  STRUCT
   GRAPHIC_INIT : BOOL ;	//NEW FL Graphic Init
   EMERGENCY_BLINK : BOOL ;	//NEW FL Emergency Blink
   ON_SW : BOOL ;	//NEW FLS On Sw Temporary
   COMPRESSED_AIR : BOOL ;	//NEW FLS Compressed Air
   AERIAL_LINK_RUN_PB : BOOL ;	//NEW FLS 508 Link Run SW - Diabled
   PACKET_in_FLIPPER_SW : BOOL ;	//NEW FLS Service Enable Switch - Disabled
   SERVICE_INIT_PB : BOOL ;	//NEW FLS Service Initialisation PB
   ALL_SERVICE_ENABLE_SW : BOOL ;	//NEW FLS All Services Enable Switch
   SERVICE_SW_1_STATUS : BOOL ;	//NEW FLS Service 1 Switch
   SERVICE_SW_2_STATUS : BOOL ;	//NEW FLS Service 2 Switch
   SERVICE_SW_3_STATUS : BOOL ;	//NEW FLS Service 3 Switch
   SERVICE_SW_1_2_STATUS : BOOL ;	//NEW FLS Service 1 or 2 Switch
   BIT12 : BOOL ;	//NEW FLS Spare
   BIT13 : BOOL ;	//NEW FLS Spare
   SERVICE_SW_2_TIME_ADJ : BOOL ;	//NEW FLS Service 2 Switch - Time Adjust
   PACKETIZER_GATE_STATUS : BOOL ;	//NEW FLS 2145 Packetizer Flap Gate - Status Bit
   E_STOP_CONSOLE_STATUS : BOOL ;	//NEW FL E-Stop Console
   E_STOP_ELEVATOR_STATUS : BOOL ;	//NEW FL E-Stop Elevator
   E_STOP_FLIPPER_STATUS : BOOL ;	//NEW FL E-Stop Flipper
   E_STOP_LOADER_STATUS : BOOL ;	//NEW FL E-Stop Loader
   HAND_FEED_ARROW_STATUS : BOOL ;	//NEW FL Hand Feed Arrow
   ELEVATOR_DOOR_STATUS : BOOL ;	//NEW FL Elevator Door
   FLIPPER_DOOR_STATUS : BOOL ;	//NEW FL Flipper Door
   LOADER_DOOR_STATUS : BOOL ;	//NEW FL Loader Door
   LIGHT_BARRIER_1_STATUS : BOOL ;	//NEW FL Light Barrier 1 - B5.4 Conveyor 1 Exit - Status Bit
   LIGHT_BARRIER_2_STATUS : BOOL ;	//NEW FL Light Barrier 2 - B5.5 Conveyor 2 InFeed - Status Bit
   LIGHT_BARRIER_3_STATUS : BOOL ;	//NEW FL Light Barrier 3 - B6.0 Conveyor 2 Presence - Status Bit
   LIGHT_BARRIER_4_STATUS : BOOL ;	//NEW FL Light Barrier 4 - B6.1 Conveyor 2 Exit - Status Bit
   LIGHT_BARRIER_5_STATUS : BOOL ;	//NEW FL Light Barrier 5 - B6.2 Conveyor 3 InFeed - Status Bit
   LIGHT_BARRIER_6_STATUS : BOOL ;	//NEW FL Light Barrier 6 - B6.4 Conveyor 3 Exit - Status Bit
   LIGHT_BARRIER_B_STATUS : BOOL ;	//NEW FL Light Barrier B - B5.2 Elevator Limit - Status Bit
   LIGHT_BARRIER_A_STATUS : BOOL ;	//NEW FL Light Barrier A - B5.1 Elevator InFeed - Status Bit
   BIT32 : BOOL ;	//NEW FL Pusher 0 Motion
   BIT33 : BOOL ;	//NEW FL Pusher 0 Motion
   BIT34 : BOOL ;	//NEW FL Pusher 0 Motion
   BIT35 : BOOL ;	//NEW FL Pusher 0 Motion
   BIT36 : BOOL ;	//NEW FL Pusher 0 Motion
   BIT37 : BOOL ;	//NEW FL Pusher 0 Motion
   BIT38 : BOOL ;	//NEW FL Pusher 0 Motion
   BIT39 : BOOL ;	//NEW FL Pusher 0 Motion
   BIT40 : BOOL ;	//NEW FL Elevator Motion
   BIT41 : BOOL ;	//NEW FL Elevator Motion
   BIT42 : BOOL ;	//NEW FL Elevator Motion
   BIT43 : BOOL ;	//NEW FL Elevator Motion
   BIT44 : BOOL ;	//NEW FL Elevator Motion
   BIT45 : BOOL ;	//NEW FL Elevator Motion
   BIT46 : BOOL ;	//NEW FL Elevator Motion
   BIT47 : BOOL ;	//NEW FL Elevator Motion
   BIT48 : BOOL ;	//NEW FL Pusher 1 Motion
   BIT49 : BOOL ;	//NEW FL Pusher 1 Motion
   BIT50 : BOOL ;	//NEW FL Pusher 1 Motion
   BIT51 : BOOL ;	//NEW FL Pusher 1 Motion
   BIT52 : BOOL ;	//NEW FL Pusher 1 Motion
   BIT53 : BOOL ;	//NEW FL Pusher 1 Motion
   BIT54 : BOOL ;	//NEW FL Pusher 1 Motion
   BIT55 : BOOL ;	//NEW FL Pusher 1 Motion
   BIT56 : BOOL ;	//NEW FL Pusher 2 Motion
   BIT57 : BOOL ;	//NEW FL Pusher 2 Motion
   BIT58 : BOOL ;	//NEW FL Pusher 2 Motion
   BIT59 : BOOL ;	//NEW FL Pusher 2 Motion
   BIT60 : BOOL ;	//NEW FL Pusher 2 Motion
   BIT61 : BOOL ;	//NEW FL Pusher 2 Motion
   BIT62 : BOOL ;	//NEW FL Pusher 2 Motion
   CONVEYORS_CLEARING : BOOL ;	//NEW FL Conveyors Clearing
   ELEVATOR_MOTOR_STATUS : BOOL ;	//NEW FL Elevator - Motor M42.0 Status Bit
   PUSHER_1_MOTOR_STATUS : BOOL ;	//NEW FL Pusher 1 - Motor M42.6 Status Bit
   CONVEYOR_1_MOTOR_STATUS : BOOL ;	//NEW FL Conv 1 - Motor M43.0 Status Bit
   CONVEYOR_2B_MOTOR_STATUS : BOOL ;	//NEW FL Conv 2 Belt - Motor M43.4 Status Bit
   CONVEYOR_2R_MOTOR_STATUS : BOOL ;	//NEW FL Conv 2 Roller - Motor M43.5 Status Bit
   CONVEYOR_3_MOTOR_STATUS : BOOL ;	//NEW FL Conveyor 3 - Motor M44.0 Status Bit
   CONVEYOR_4_MOTOR_STATUS : BOOL ;	//NEW FL Conveyor 4 - Motor M44.3 Status Bit
   CONVEYOR_5_MOTOR_STATUS : BOOL ;	//NEW FL Conveyor 5 - Motor M45.0 Status Bit
   CONVEYOR_6_MOTOR_STATUS : BOOL ;	//NEW FL Conveyor 6 - Motor M45.3 Status Bit
   CONVEYOR_7_MOTOR_STATUS : BOOL ;	//NEW FL Conveyor 7 - Motor M45.6 Status Bit
   FLIPPER_MOTOR_STATUS : BOOL ;	//NEW FL Flipper Flip - Motor M46.0 Status Bit
   CONVEYOR_8_MOTOR_STATUS : BOOL ;	//NEW FL Conveyor 8 - Motor M46.4 Status Bit
   TURNTABLE_MOTOR_STATUS : BOOL ;	//NEW FL TurnTable - Motor M47.0 Status Bit
   CONVEYOR_9_MOTOR_STATUS : BOOL ;	//NEW FL Conveyor 9 - Motor M47.5 Status Bit
   PUSHER_2_MOTOR_STATUS : BOOL ;	//NEW FL Pusher 2 - Motor M47.6 Status Bit
   CONVEYOR_10_MOTOR_STATUS : BOOL ;	//NEW FL Conveyor 10 - Motor M48.0 Status Bit
   CONVEYOR_11_MOTOR_STATUS : BOOL ;	//NEW FL Conveyor 11 - Motor M48.3 Status Bit
   CONVEYOR_12_MOTOR_STATUS : BOOL ;	//NEW FL Conveyor 12 - Motor M48.6 Status Bit
   CONVEYOR_13_MOTOR_STATUS : BOOL ;	//NEW FL Conveyor 13 - Motor M49.0 Status Bit
   CONVEYOR_21_MOTOR_STATUS : BOOL ;	//NEW FL Conveyor 21 - Motor M53.2 Status Bit
   CONVEYOR_22_MOTOR_STATUS : BOOL ;	//NEW FL Conveyor 22 - Motor M53.4 Status Bit
   CONVEYOR_23_MOTOR_STATUS : BOOL ;	//NEW FL Conveyor 23 - Motor M54.0 Status Bit
   LOADER_LIFT_MOTOR_STATUS : BOOL ;	//NEW FL Loader Lift - Motor M50.0 Status Bit
   LOADER_FING_MOTOR_STATUS : BOOL ;	//NEW FL Loader Fingers - Motor M50.5 Status Bit
   LOADER_BELT_MOTOR_STATUS : BOOL ;	//NEW FL Loader Belt - Motor M51.0 Status Bit
   LIGHT_BARRIER_7_STATUS : BOOL ;	//NEW FL Light Barrier 7 - B6.7 Conv 4 InFeed Sens - Status
   LIGHT_BARRIER_8_STATUS : BOOL ;	//NEW FL Light Barrier 8 - B7.0 Conv 4 Exit Sens - Status
   LIGHT_BARRIER_9_STATUS : BOOL ;	//NEW FL Light Barrier 9 - B7.1 Conv 5 Exit Sens - Status
   LIGHT_BARRIER_10_STATUS : BOOL ;	//NEW FL Light Barrier 10 - B7.2 Conv 6 Slow Sens - Status Bit
   LIGHT_BARRIER_11_STATUS : BOOL ;	//NEW FL Light Barrier 11 - B7.3 Conv 6 Exit Sens - Status Bit
   LIGHT_BARRIER_12_STATUS : BOOL ;	//NEW FL Light Barrier 12 - B7.4 FLipper InFeed Sens - Status Bit
   LIGHT_BARRIER_13_STATUS : BOOL ;	//NEW FL Light Barrier 13 - B8.2 Flipper Exit Sens - Status Bit
   LIGHT_BARRIER_14_STATUS : BOOL ;	//NEW FL Light Barrier 14 - B9.6 Conv 9 InFeed Sens - Status Bit
   LIGHT_BARRIER_15_STATUS : BOOL ;	//NEW FL Light Barrier 15 - B9.7 Conv 9 Packet Sens - Status Bit
   LIGHT_BARRIER_16_STATUS : BOOL ;	//NEW FL Light Barrier 16 - B10.3 Conv 10 Start Sens - Status Bit
   LIGHT_BARRIER_17_STATUS : BOOL ;	//NEW FL Light Barrier 17 - B10.4 Conv 10 InFeed Sens - Status Bit
   LIGHT_BARRIER_18_STATUS : BOOL ;	//NEW FL Light Barrier 18 - B10.5 Conv 10 Full Sens - Status Bit
   LIGHT_BARRIER_19_STATUS : BOOL ;	//NEW FL Light Barrier 19 - B10.6 Conv 10 Exit Sens - Status Bit
   LIGHT_BARRIER_20_STATUS : BOOL ;	//NEW FL Light Barrier 20 - B10.7 Conv 11 Exit Sens - Status Bit
   LIGHT_BARRIER_21_STATUS : BOOL ;	//NEW FL Light Barrier 21 - B11.0 Conv 12 Exit Sens - Status Bit- Status Bit
   LIGHT_BARRIER_22_STATUS : BOOL ;	//NEW FL Light Barrier 22 - B11.1 Conv 13 Slow Sens - Status Bit
   LIGHT_BARRIER_23_STATUS : BOOL ;	//NEW FL Light Barrier 23 - B11.2 Conv 13 Exit Sens - Status Bit
   LIGHT_BARRIER_24_STATUS : BOOL ;	//NEW FL Light Barrier 24 - B12.3 Fingers Delivery Sens - Status Bit
   LIGHT_BARRIER_25_STATUS : BOOL ;	//NEW FL Light Barrier 25 - B13.0 Loader Empty Sens - Status Bit
   LIGHT_BARRIER_26_STATUS : BOOL ;	//NEW FL Light Barrier 26 - B15.4 Conv 21 Exit Sens - Status Bit
   LIGHT_BARRIER_27_STATUS : BOOL ;	//NEW FL Light Barrier 27 - B15.5 Conv 22 Exit Sens - Status Bit
   LIGHT_BARRIER_28_STATUS : BOOL ;	//NEW FL Light Barrier 28 - B15.6 Conv 23 Slow Sens - Status Bit
   LIGHT_BARRIER_29_STATUS : BOOL ;	//NEW FL Light Barrier 29 - B15.7 Conv 23 Exit Sens - Status Bit
   LIGHT_BARRIER_30_STATUS : BOOL ;	//NEW FL Light Barrier 30 - B35.2 Conv 0 InFeed Sens - Status Bit
   LIGHT_BARRIER_31_STATUS : BOOL ;	//NEW FL Light Barrier 31 - B35.3 Conv 0 Exit Sens - Status Bit
   LIGHT_BARRIER_32_STATUS : BOOL ;	//NEW FL Light Barrier 32 - B35.4 Conv 0 Length Sens - Status Bit
   PROX_9_STATUS : BOOL ;	//NEW FL Prox 9 - P8.5 TurnTable Rotation InFeed Slow - Status Bit
   PROX_10_STATUS : BOOL ;	//NEW FL Prox 10 - P8.6 TurnTable Rotation InFeed Stop - Status Bit
   PROX_11_STATUS : BOOL ;	//NEW FL Prox 11 - P9.2 TurnTable Rotation Exit Slow - Status Bit
   PROX_12_STATUS : BOOL ;	//NEW FL Prox 12 - P9.3 TurnTable Rotation Exit Stop - Status Bit
   PROX_13_STATUS : BOOL ;	//NEW FL Prox 13 - P10.0 Pusher 2 Retract Sens - Status Bit
   PROX_14_STATUS : BOOL ;	//NEW FL Prox 14 - P10.1 Pusher 2 Extend Sens - Status Bit
   PROX_15_STATUS : BOOL ;	//NEW FL Prox 15 - P15.0 Pivot 10 High Sens - Status Bit
   PROX_16_STATUS : BOOL ;	//NEW FL Prox 16 - P15.1 Pivot 10 Low Sens - Status Bit
   PROX_17_STATUS : BOOL ;	//NEW FL Prox 17 - P13.2 Loader H Level Stop - Status Bit
   PROX_18_STATUS : BOOL ;	//NEW FL Prox 18 - P13.1 Loader H Level Slow - Status Bit
   PROX_19_STATUS : BOOL ;	//NEW FL Prox 19 - P11.4 Loader L Level Stop - Status Bit
   PROX_20_STATUS : BOOL ;	//NEW FL Prox 20 - P11.5 Loader L Level Slow - Status Bit
   PROX_21_STATUS : BOOL ;	//NEW FL Prox 21 - P11.6 Loader Slow Bot - Status Bit
   PROX_22_STATUS : BOOL ;	//NEW FL Prox 22 - P11.7 Loader Stop Bot - Status Bit
   PROX_23_STATUS : BOOL ;	//NEW FL Prox 23 - P12.0 Loader Finger Retract - Status Bit
   PROX_24_STATUS : BOOL ;	//NEW FL Prox 24 - P12.1 Loader Finger Extend - Status Bit
   FP131 : BOOL ;	//NEW FP One Shot
   FP132 : BOOL ;	//NEW FP One Shot
   FP133 : BOOL ;	//NEW FP One Shot
   FP134 : BOOL ;	//NEW FP One Shot
   FP135 : BOOL ;	//NEW FP One Shot
   TURNTABLE_DELIV_POSITION : BOOL ;	//NEW FL TurnTable Delivery Position
   TURNTABLE_REVERSE_ARROW : BOOL ;	//NEW FL TurnTable Arrow Reverse Packet
   TURNTABLE_DIR_SELECT_SW : BOOL ;	//NEW FL TurnTable Direction Select SW
   TURNTABLE_FLICK_MOTION : BOOL ;	//NEW FL TurnTable Flicker - Motion
   FP140 : BOOL ;	//NEW FP One Shot
   FP141 : BOOL ;	//NEW FP One Shot
   FP142 : BOOL ;	//NEW FP One Shot
   FP143 : BOOL ;	//NEW FP One Shot
   PROX_1_STATUS : BOOL ;	//NEW FL Prox 1 - P4.0 Elevator Bottom Position - Status Bit
   PROX_2_STATUS : BOOL ;	//NEW FL Prox 2 - P4.1 Elevator SlowDown Bot - Status Bit
   PROX_3_STATUS : BOOL ;	//NEW FL Prox 3 - P4.2 Elevator SlowDown Top - Status Bit
   PROX_4_STATUS : BOOL ;	//NEW FL Prox 4 - P4.3 Elevator Top Position - Status Bit
   PROX_5_STATUS : BOOL ;	//NEW FL Prox 5 - P4.4 Pusher 1 Home - Status Bit
   PROX_6_STATUS : BOOL ;	//NEW FL Prox 6 - P4.5 Pusher 1 Limit - Status Bit
   PROX_7_STATUS : BOOL ;	//NEW FL Prox 7 - P8.0 Flipper Fingers Right Position - Status Bit
   PROX_8_STATUS : BOOL ;	//NEW FL Prox 8 - P8.1 Flipper Fingers Left Position - Status Bit
   BIT152 : BOOL ;	//NEW FL Loader Motion
   BIT153 : BOOL ;	//NEW FL Loader Motion
   BIT154 : BOOL ;	//NEW FL Loader Motion
   BIT155 : BOOL ;	//NEW FL Loader Motion
   BIT156 : BOOL ;	//NEW FL Loader Motion
   BIT157 : BOOL ;	//NEW FL Loader Motion
   BIT158 : BOOL ;	//NEW FL Loader Motion
   BIT159 : BOOL ;	//NEW FL Loader Motion
   SERVICE_SSW_MAIN : BOOL ;	//NEW FL Service SW Main Screen
   SERVICE_SSW_STATUS : BOOL ;	//NEW FL Service SW Main Screen - Status
   CLEARING_SSW_MAIN : BOOL ;	//NEW FL Clearing SW Main Screen
   CLEARING_SSW_STATUS : BOOL ;	//NEW FL Clearing SW Main Screen - Status
   MAN_FEED_SSW_MAIN : BOOL ;	//NEW FL Hand Feed SW Main Screen
   MAN_FEED_SSW_STATUS : BOOL ;	//NEW FL Hand Feed SW Main Screen - Status
   TURNTABLE_SSW_MAIN : BOOL ;	//NEW FL Turn Table Turn SW = 1:CCW - 0:CW Main Screen
   TURNTABLE_SSW_STATUS : BOOL ;	//NEW FL Turn Table Select Main Screen - Status
   FLIPPER_SSW_MAIN : BOOL ;	//NEW FL Flipper SW Main Screen
   FLIPPER_SSW_STATUS : BOOL ;	//NEW FL Flipper SW Main Screen - Status
   ROLLER_SSW_MAIN : BOOL ;	//NEW FL Roller SW Main Screen
   ROLLER_SSW_STATUS : BOOL ;	//NEW FL Roller SW Main Screen - Status
   ELEVATOR_ROUND_TRIP_SSW : BOOL ;	//NEW FL Elevator - Round Trip PB
   BIT173 : BOOL ;
   BIT174 : BOOL ;
   BIT175 : BOOL ;
   HMI_PUSHER_0_TEST_SSW : BOOL ;	//NEW FL Pusher 0 SW
   HMI_ELEVATOR_SERVICE_SSW : BOOL ;	//NEW FL Elevator Service SW
   HMI_ELEVATOR_TEST_DN_SSW : BOOL ;	//NEW FL Elevator DN PB
   HMI_ELEVATOR_TEST_UP_SSW : BOOL ;	//NEW FL Elevator UP PB
   HMI_ROLLER_TEST_FWD_SSW : BOOL ;	//NEW FL Roller FWD SW
   HMI_ROLLER_TEST_REV_SSW : BOOL ;	//NEW FL Roller REV SW
   HMI_PUSHER_1_TEST_SSW : BOOL ;	//NEW FL Pusher 1 SW
   HMI_CONVEYOR_1_TEST_SSW : BOOL ;	//NEW FL Conv 1 SW
   HMI_CONVEYOR_2B_TEST_SSW : BOOL ;	//NEW FL Conv 2 Belt SW
   HMI_CONVEYOR_2L_TEST_SSW : BOOL ;	//NEW FL Conv 2 Lift SW
   HMI_CONVEYOR_2R_TEST_SSW : BOOL ;	//NEW FL Conv 2 Roller SW
   HMI_CONVEYOR_3_TEST_SSW : BOOL ;	//NEW FL Conv 3 SW
   HMI_CONVEYOR_4_TEST_SSW : BOOL ;	//NEW FL Conv 4 SW
   HMI_CONVEYOR_5_TEST_SSW : BOOL ;	//NEW FL Conv 5 SW
   HMI_CONVEYOR_6_TEST_SSW : BOOL ;	//NEW FL Conv 6 SW
   HMI_CONVEYOR_7_TEST_SSW : BOOL ;	//NEW FL Flipper Conv 7 SW
   HMI_CONVEYOR_8_TEST_SSW : BOOL ;	//NEW FL Turn Table Conv 8 SW
   HMI_TURNTABLE_CCW_SSW : BOOL ;	//NEW FL Turn Table / Conveyor CCW PB
   HMI_TURNTABLE_CW_SSW : BOOL ;	//NEW FL Turn Table / Conveyor CW PB
   HMI_FLIPPER_SERVICE_SSW : BOOL ;	//NEW FL Flipper Service SW
   HMI_FLIPPER_FLIP_SSW : BOOL ;	//NEW FL Flipper - Flip PB
   HMI_CONVEYOR_9_TEST_SSW : BOOL ;	//NEW FL Conv 9 SW
   HMI_PUSHER_2_TEST_SSW : BOOL ;	//NEW FL Pusher 2 SW
   HMI_PIVOT_SERVICE_SSW : BOOL ;	//NEW FL Conv 10 - Pivot Service SW
   HMI_PIVOT_TEST_DN_SSW : BOOL ;	//NEW FL Conv 10 - Pivot DN PB
   HMI_PIVOT_TEST_UP_SSW : BOOL ;	//NEW FL Conv 10 - Pivot UP PB
   BIT202 : BOOL ;	//NEW FL Spare
   BIT203 : BOOL ;	//NEW FL Spare
   TURNTABLE_SERVICE_PBSHOW : BOOL ;	//NEW FL TurnTable Service PB SHOW
   TURNTABLE_SERVICE_SSW : BOOL ;	//NEW FL TurnTable Service SW
   HMI_CONVEYOR_10_TEST_SSW : BOOL ;	//NEW FL Conv 10 - Conveyor SW
   LOADER_FING_SERVICE_SSW : BOOL ;	//NEW FL Loader Service SW - Fingers
   LOADER_LIFT_SERVICE_SSW : BOOL ;	//NEW FL Loader Service SW - Lift
   LOADER_LIFT_TOP_PB : BOOL ;	//NEW FL Loader Lift - TOP PB
   LOADER_LIFT_UP_PB : BOOL ;	//NEW FL Loader Lift - UP PB
   LOADER_LIFT_DN_PB : BOOL ;	//NEW FL Loader Lift - DOWN PB
   FINGER_RETRACT_TEST_PB : BOOL ;	//NEW FL Loader Fingers Retract PB
   FINGER_EXTEND_TEST_PB : BOOL ;	//NEW FL Loader Fingers Extend PB
   FINGER_TILT_TEST_PB : BOOL ;	//NEW FL Loader Fingers Tilt Down PB
   FINGER_BELT_TEST_SW : BOOL ;	//NEW FL Loader Fingers Belt SW
   HMI_CONVEYOR_11_TEST_SSW : BOOL ;	//NEW FL Conv 11 Test SW
   HMI_CONVEYOR_12_TEST_SSW : BOOL ;	//NEW FL Conv 12 Test SW
   HMI_CONVEYOR_13_TEST_SSW : BOOL ;	//NEW FL Conv 13 Test SW
   HMI_CONVEYOR_21_TEST_SSW : BOOL ;	//NEW FL Conv 21 Test SW
   HMI_CONVEYOR_22_TEST_SSW : BOOL ;	//NEW FL Conv 22 Test SW
   HMI_CONVEYOR_23_TEST_SSW : BOOL ;	//NEW FL Conv 23 Test SW
   CONVEYOR_0_MOTOR_STATUS : BOOL ;	//NEW FL Conveyor 0 - Motor M62.0 Status Bit
   PUSHER_0_MOTOR_STATUS : BOOL ;	//NEW FL Pusher 0 - Motor M62.2 Status Bit
   PUSHER_0_COLOR_WORD : WORD ;	//NEW WD Pusher 0 - 2145 - Motor Status Color
   CONV_0_COLOR_WORD : WORD ;	//NEW WD Conveyor 0 - 2145 - Motor Status Color
   ELEVATOR_COLOR_WORD : WORD ;	//NEW WD Elevator - Motor Status Color
   PUSHER_1_COLOR_WORD : WORD ;	//NEW WD Pusher 1 - Motor Status Color
   CONV_1_COLOR_WORD : WORD ;	//NEW WD Conv 1 - Motor Status Color
   CONV_2_BELT_COLOR_WORD : WORD ;	//NEW WD Conv 2 Belt - Motor Status Color
   LIFT_ROLLER_2_COLOR_WORD : WORD ;	//NEW WD Lift 2 Roller - Actuator Status Color
   CONV_2_ROLLER_COLOR_WORD : WORD ;	//NEW WD Conv 2 Roller - Motor Status Color
   CONV_3_COLOR_WORD : WORD ;	//NEW WD Conveyor 3 - Motor Status Color
   CONV_4_COLOR_WORD : WORD ;	//NEW WD Conveyor 4 - Motor Status Color
   CONV_5_COLOR_WORD : WORD ;	//NEW WD Conveyor 5 - Motor Status Color
   CONV_6_COLOR_WORD : WORD ;	//NEW WD Conveyor 6 - Motor Status Color
   CONV_7_COLOR_WORD : WORD ;	//NEW WD Conveyor 7 - Motor Status Color
   FLIPPER_COLOR_WORD : WORD ;	//NEW WD Flipper - Motor M46.0 Status Color
   CONV_8_COLOR_WORD : WORD ;	//NEW WD Conveyor 8 - Motor M46.4 Status Color
   TURN_TABLE_COLOR_WORD : WORD ;	//NEW WD TurnTable - Motor M47.0 Status Color
   CONV_9_COLOR_WORD : WORD ;	//NEW WD Conveyor 9 - Motor M47.5 Status Color
   PUSHER_2_COLOR_WORD : WORD ;	//NEW WD Pusher 2 - Motor M47.6 Status Color
   CONV_10_COLOR_WORD : WORD ;	//NEW WD Conveyor 10 - Motor M48.0 Status Color
   CONV_11_COLOR_WORD : WORD ;	//NEW WD Conveyor 11 - Motor M48.3 Status Color
   CONV_12_COLOR_WORD : WORD ;	//NEW WD Conveyor 12 - Motor M48.6 Status Color
   CONV_13_COLOR_WORD : WORD ;	//NEW WD Conveyor 13 - Motor M49.0 Status Color
   CONV_21_COLOR_WORD : WORD ;	//NEW WD Conveyor 21 - Motor M53.4 Status Color
   CONV_22_COLOR_WORD : WORD ;	//NEW WD Conveyor 22 - Motor M53.6 Status Color
   CONV_23_COLOR_WORD : WORD ;	//NEW WD Conveyor 23 - Motor M54.0 Status Color
   LOADER_LIFT_COLOR_WORD : WORD ;	//NEW WD Loader Lift - Motor M54.6 Status Color
   LOADER_FING_COLOR_WORD : WORD ;	//NEW WD Loader Fingers - Motor M50.5 Status Color
   FINGERS_BELT_COLOR_WORD : WORD ;	//NEW WD Fingers Belt - Motor M54.6 Status Color
   HIGH_LEVEL_23_GRAPHIC : WORD ;	//NEW WD High Level Conveyor 23
   LOW_LEVEL_13_GRAPHIC : WORD ;	//NEW WD Low Level Conveyor 13
   PIVOT_GRAPHIC : WORD ;	//NEW WD Pivot Conveyor Graphic
   CONV_3_COUNT : WORD ;	//NEW WD Slat Conveyor 3 - Packet Count
   CONV_4_COUNT : WORD ;	//NEW WD Collator Conveyor 4 - Packet Count
   CONV_5_COUNT : WORD ;	//NEW WD Link Conveyor 5 - Packet Count
   CONV_6_COUNT : WORD ;	//NEW WD Delivery Conveyor 6 - Packet Count
   CONV_10_COUNT : WORD ;	//NEW WD Pivot Conveyor 10 - Packet Count
   CONV_11_COUNT : WORD ;	//NEW WD Cumul Conveyor 11 - Packet Count
   CONV_12_COUNT : WORD ;	//NEW WD Cumul Conveyor 12 - Packet Count
   CONV_13_COUNT : WORD ;	//NEW WD Delivery Conveyor 13 - Packet Count
   CONV_21_COUNT : WORD ;	//NEW WD Cumul Conveyor 21 - Packet Count
   CONV_22_COUNT : WORD ;	//NEW WD Cumul Conveyor 22 - Packet Count
   CONV_23_COUNT : WORD ;	//NEW WD Delivery Conveyor 23 - Packet Count
   FLIPPER_CCW : WORD ;	//NEW WD Flipper Graphic CCW
   FLIPPER_CW : WORD ;	//NEW WD Flipper Graphic CW
   FLIPPER_POSITION : WORD ;	//NEW WD Flipper Positioning mS
   TURN_COLOR : WORD ;	//NEW WD Turn Table - Turn Color
   FLIPPER_COLOR : WORD ;	//NEW WD Flipper Color
   FLIPPER_PACK_PRESENCE : WORD ;	//NEW WD Flipper - Packet Presence
   TURNTABLE_PACK_PRESENCE : WORD ;	//NEW WD TurnTable - Packet Presence
   ROLLER_PACK_PRESENCE : WORD ;	//NEW WD Pusher Roller - Packet Presence
   PUSHER_PACK_PRESENCE : WORD ;	//NEW WD Pusher - Packet Presence
   CONV_0_STATUS : BOOL ;	//NEW FL Conveyor 0 - Motor Status Bit
   PUSHER_0_STATUS : BOOL ;	//NEW FL Pusher 0 - Motor Status
   ELEVATOR_STATUS : BOOL ;	//NEW FL Elevator - Motor Status
   PUSHER_1_STATUS : BOOL ;	//NEW FL Pusher 1 - Motor Status
   CONV_1_STATUS : BOOL ;	//NEW FL Conveyor 1 - Motor Status
   TURNTABLE_RNDTRIP : BOOL ;	//NEW FL TurnTable Round Trip CMD
   RNDTRIP_PB_VISIBLE : BOOL ;	//NEW FL TurnTable Round Trip PB Visible
   BOOL_SPARE227 : BOOL ;	//NEW FL
   SCREEN_CALL_0 : BOOL ;	//NEW FL  HMI Call Screen 0
   SCREEN_CALL_1 : BOOL ;	//NEW FL  HMI Call Screen 1
   SCREEN_CALL_2 : BOOL ;	//NEW FL  HMI Call Screen 2
   SCREEN_CALL_3 : BOOL ;	//NEW FL  HMI Call Screen 3
   SCREEN_CALL_4 : BOOL ;	//NEW FL  HMI Call Screen 4
   BOOL_SPARE2276 : BOOL ;	//NEW FL
   BOOL_SPARE2277 : BOOL ;	//NEW FL
   BOOL_SPARE2278 : BOOL ;	//NEW FL
   BOOL_SPARE2279 : BOOL ;	//NEW FL
   BOOL_SPARE22710 : BOOL ;	//NEW FL
   BOOL_SPARE22711 : BOOL ;	//NEW FL
   BOOL_SPARE22712 : BOOL ;	//NEW FL
   BOOL_SPARE22713 : BOOL ;	//NEW FL
   BOOL_SPARE22714 : BOOL ;	//NEW FL
   BOOL_SPARE22715 : BOOL ;	//NEW FL
   BOOL_SPARE22716 : BOOL ;	//NEW FL
   BOOL_SPARE22717 : BOOL ;	//NEW FL
   BOOL_SPARE22718 : BOOL ;	//NEW FL
   BOOL_SPARE22719 : BOOL ;	//NEW FL
   BOOL_SPARE22720 : BOOL ;	//NEW FL
   BOOL_SPARE22721 : BOOL ;	//NEW FL
   BOOL_SPARE22722 : BOOL ;	//NEW FL
   BOOL_SPARE22723 : BOOL ;	//NEW FL
   BOOL_SPARE22724 : BOOL ;	//NEW FL
   WORD_SPARE23 : WORD ;	//NEW WD
   FLIPPER_TURN_COLOR : WORD ;	//NEW WD Flipper Turn Color
   NEW_ORDER_COLOR : WORD ;	//NEW WD Conveyor 10 - New Order Color
   SERVICE_FLIPPER : BOOL ;	//NEW FLS Flipper Service - Switch
   FLIP_TEST : BOOL ;	//NEW FLS Flipper Flip - Test Switch
   SERVICE_TURNTABLE : BOOL ;	//NEW FLS TurnTable Service - Switch
   TURN_TEST_CW : BOOL ;	//NEW FLS TurnTable - Turn CW - Status Bit
   TURN_TEST_CCW : BOOL ;	//NEW FLS TurnTable - Turn CCW - Status Bit
   PUSHER_2_TEST : BOOL ;	//NEW FLS Pusher 2 - Test Switch
   CONVEYOR_10_TEST_SW : BOOL ;	//NEW FLS Collator Conveyor 10 - Test Switch
   PIVOT_SERVICE_SW : BOOL ;	//NEW FL Pivot Service - Status
   PIVOT_UP_TEST_PB : BOOL ;	//NEW FLS Pivot Conveyor UP - Test Switch
   PIVOT_DN_TEST_PB : BOOL ;	//NEW FLS Pivot Conveyor DN - Test Switch
   PIVOT_STATUS : BOOL ;	//NEW FL Pivot ON - Status
   CONV_8_INVERT_SELECT : BOOL ;	//NEW FL TurnTable Conveyor 8 - Positioning Time - Display Selector Bit - INVERT
   CONVEYOR_11_TEST_SW : BOOL ;	//NEW FLS Cumul Conveyor 11 - Test Switch
   CONVEYOR_12_TEST_SW : BOOL ;	//NEW FLS Cumul Conveyor 12 - Test Switch
   CONVEYOR_13_TEST_SW : BOOL ;	//NEW FLS Delivery Conveyor 13 - Test Switch
   CONVEYOR_21_TEST_SW : BOOL ;	//NEW FLS Cumul Conveyor 21 - Test Switch
   CONVEYOR_22_TEST_SW : BOOL ;	//NEW FLS Cumul Conveyor 22 - Test Switch
   CONVEYOR_23_TEST_SW : BOOL ;	//NEW FLS Delivery Conveyor 23 - Test Switch
   LOADER_SERVICE_SW : BOOL ;	//NEW FLS Loader Service - Switch
   LOADER_UP_TEST_PB : BOOL ;	//NEW FLS Loader Lift Up - Test Switch
   LOADER_DN_TEST_PB : BOOL ;	//NEW FLS Loader Lift Dn - Test Switch
   FINGERS_EXTEND_TEST_PB : BOOL ;	//NEW FLS Loader Finger Extend - Test Switch
   FINGERS_RETRACT_TEST_PB : BOOL ;	//NEW FLS Loader Finger Retract - Test Switch
   FP_ONESHOT_0 : BOOL ;	//NEW FP One Shot
   CONVEYOR_0_SERVICE_SW : BOOL ;	//NEW FL Conveyor 0 / Pusher 0 - Service Enable
   ELEVATOR_SERVICE_SW : BOOL ;	//NEW FL Elevator / Pusher 1 - Service Enable
   CONVEYOR_1_SERVICE_SW : BOOL ;	//NEW FL Conveyor 1 - Service Enable Select - Screen 4
   CONVEYOR_2_SERVICE_SW : BOOL ;	//NEW FL Conveyor 2 - Service Enable Select - Screen 4
   CONVEYOR_3_SERVICE_SW : BOOL ;	//NEW FL Conveyor 3 - Service Enable Select - Screen 4
   CONVEYOR_4_SERVICE_SW : BOOL ;	//NEW FL Conveyor 4 - Service Enable Select - Screen 4
   CONVEYOR_5_SERVICE_SW : BOOL ;	//NEW FL Conveyor 5 - Service Enable Select - Screen 4
   CONVEYOR_6_SERVICE_SW : BOOL ;	//NEW FL Conveyor 6 - Service Enable Select - Screen 4
   CONVEYOR_7_SERVICE_SW : BOOL ;	//NEW FL Conveyor 7 / Flipper - Service Enable Select - Screen 4
   CONVEYOR_8_SERVICE_SW : BOOL ;	//NEW FL Conveyor 8 / TurnTable - Service Enable Select - Screen 4
   CONVEYOR_9_SERVICE_SW : BOOL ;	//NEW FL Conveyor 9 / Pusher 2 - Service Enable Select - Screen 4
   CONVEYOR_10_SERVICE_SW : BOOL ;	//NEW FL Conveyor 10 - Service Enable Select - Screen 4
   CONVEYOR_11_SERVICE_SW : BOOL ;	//NEW FL Conveyors 11, 12, 13 - Service Enable Select - Screen 4
   CONVEYOR_21_SERVICE_SW : BOOL ;	//NEW FL Conveyors 21, 22, 23 - Service Enable Select - Screen 4
   LOADER_SERVICE_ENABLE_SW : BOOL ;	//NEW FL Loader - Service Enable
   CTRL48 : BOOL ;	//NEW FL Spare - Service Enable
   CTRL49 : BOOL ;	//NEW FL Spare -
   CTRL50 : BOOL ;	//NEW FL Spare -
   CTRL51 : BOOL ;	//NEW FL Spare -
   CTRL52 : BOOL ;	//NEW FL Spare -
   CTRL53 : BOOL ;	//NEW FL Spare -
   CTRL54 : BOOL ;	//NEW FL Spare -
   CTRL55 : BOOL ;	//NEW FL Spare -
   CTRL56 : BOOL ;	//NEW FL Spare -
   CLEARING_FUNCTION : WORD ;	//NEW WD Clearing Function - Underneat Rectangle
   WORD57 : WORD ;	//NEW WD
   WORD58 : WORD ;	//NEW WD
   ACTUAL_HMI_SCREEN_NO : WORD ;	//NEW WD HMI Actual Display Screen
   CONVEYOR_MAXCOUNT_L : WORD  := W#16#6;	//NEW WD All Conveyors Max Count Lenght (6)
   CONVEYOR_MAXCOUNT_W : WORD  := W#16#7;	//NEW WD All Conveyors Max Count Widtht (7)
   WORD62 : WORD ;	//NEW WD
   CONV_7_POS_mS : WORD ;	//NEW WD Flipper Conveyor 7 - Positioning Time x10 [mS]
   CONV_8_POS_FWD_mS : WORD ;	//NEW WD TurnTable Conveyor 8 - FWD Positioning Time x10 [mS]
   CONV_8_POS_REV_mS : WORD ;	//NEW WD TurnTable Conveyor 8 - REV Positioning Time x10 [mS]
   CONV_9_POS_mS : WORD ;	//NEW WD Pusher 2 Conveyor 9 - Positioning Time x10 [mS]
   WORD_PACKET_LENGTH : WORD ;	//NEW WD Actual Packet Length mm
   DELAY_DISPLAY_7 : WORD ;	//NEW WD HMI Flipper 7 Delay Display
   DELAY_DISPLAY_9 : WORD ;	//NEW WD HMI Conveyor 9 Delay Display
   WORD_SPARE2 : WORD ;
   WORD_SPARE3 : WORD ;
   WORD_SPARE4 : WORD ;
  END_STRUCT ;
BEGIN
   GRAPHIC_INIT := FALSE;
   EMERGENCY_BLINK := FALSE;
   ON_SW := FALSE;
   COMPRESSED_AIR := FALSE;
   AERIAL_LINK_RUN_PB := FALSE;
   PACKET_in_FLIPPER_SW := FALSE;
   SERVICE_INIT_PB := FALSE;
   ALL_SERVICE_ENABLE_SW := FALSE;
   SERVICE_SW_1_STATUS := FALSE;
   SERVICE_SW_2_STATUS := FALSE;
   SERVICE_SW_3_STATUS := FALSE;
   SERVICE_SW_1_2_STATUS := FALSE;
   BIT12 := FALSE;
   BIT13 := FALSE;
   SERVICE_SW_2_TIME_ADJ := FALSE;
   PACKETIZER_GATE_STATUS := FALSE;
   E_STOP_CONSOLE_STATUS := FALSE;
   E_STOP_ELEVATOR_STATUS := FALSE;
   E_STOP_FLIPPER_STATUS := FALSE;
   E_STOP_LOADER_STATUS := FALSE;
   HAND_FEED_ARROW_STATUS := FALSE;
   ELEVATOR_DOOR_STATUS := FALSE;
   FLIPPER_DOOR_STATUS := FALSE;
   LOADER_DOOR_STATUS := FALSE;
   LIGHT_BARRIER_1_STATUS := FALSE;
   LIGHT_BARRIER_2_STATUS := FALSE;
   LIGHT_BARRIER_3_STATUS := FALSE;
   LIGHT_BARRIER_4_STATUS := FALSE;
   LIGHT_BARRIER_5_STATUS := FALSE;
   LIGHT_BARRIER_6_STATUS := FALSE;
   LIGHT_BARRIER_B_STATUS := FALSE;
   LIGHT_BARRIER_A_STATUS := FALSE;
   BIT32 := FALSE;
   BIT33 := FALSE;
   BIT34 := FALSE;
   BIT35 := FALSE;
   BIT36 := FALSE;
   BIT37 := FALSE;
   BIT38 := FALSE;
   BIT39 := FALSE;
   BIT40 := FALSE;
   BIT41 := FALSE;
   BIT42 := FALSE;
   BIT43 := FALSE;
   BIT44 := FALSE;
   BIT45 := FALSE;
   BIT46 := FALSE;
   BIT47 := FALSE;
   BIT48 := FALSE;
   BIT49 := FALSE;
   BIT50 := FALSE;
   BIT51 := FALSE;
   BIT52 := FALSE;
   BIT53 := FALSE;
   BIT54 := FALSE;
   BIT55 := FALSE;
   BIT56 := FALSE;
   BIT57 := FALSE;
   BIT58 := FALSE;
   BIT59 := FALSE;
   BIT60 := FALSE;
   BIT61 := FALSE;
   BIT62 := FALSE;
   CONVEYORS_CLEARING := FALSE;
   ELEVATOR_MOTOR_STATUS := FALSE;
   PUSHER_1_MOTOR_STATUS := FALSE;
   CONVEYOR_1_MOTOR_STATUS := FALSE;
   CONVEYOR_2B_MOTOR_STATUS := FALSE;
   CONVEYOR_2R_MOTOR_STATUS := FALSE;
   CONVEYOR_3_MOTOR_STATUS := FALSE;
   CONVEYOR_4_MOTOR_STATUS := FALSE;
   CONVEYOR_5_MOTOR_STATUS := FALSE;
   CONVEYOR_6_MOTOR_STATUS := FALSE;
   CONVEYOR_7_MOTOR_STATUS := FALSE;
   FLIPPER_MOTOR_STATUS := FALSE;
   CONVEYOR_8_MOTOR_STATUS := FALSE;
   TURNTABLE_MOTOR_STATUS := FALSE;
   CONVEYOR_9_MOTOR_STATUS := FALSE;
   PUSHER_2_MOTOR_STATUS := FALSE;
   CONVEYOR_10_MOTOR_STATUS := FALSE;
   CONVEYOR_11_MOTOR_STATUS := FALSE;
   CONVEYOR_12_MOTOR_STATUS := FALSE;
   CONVEYOR_13_MOTOR_STATUS := FALSE;
   CONVEYOR_21_MOTOR_STATUS := FALSE;
   CONVEYOR_22_MOTOR_STATUS := FALSE;
   CONVEYOR_23_MOTOR_STATUS := FALSE;
   LOADER_LIFT_MOTOR_STATUS := FALSE;
   LOADER_FING_MOTOR_STATUS := FALSE;
   LOADER_BELT_MOTOR_STATUS := FALSE;
   LIGHT_BARRIER_7_STATUS := FALSE;
   LIGHT_BARRIER_8_STATUS := FALSE;
   LIGHT_BARRIER_9_STATUS := FALSE;
   LIGHT_BARRIER_10_STATUS := FALSE;
   LIGHT_BARRIER_11_STATUS := FALSE;
   LIGHT_BARRIER_12_STATUS := FALSE;
   LIGHT_BARRIER_13_STATUS := FALSE;
   LIGHT_BARRIER_14_STATUS := FALSE;
   LIGHT_BARRIER_15_STATUS := FALSE;
   LIGHT_BARRIER_16_STATUS := FALSE;
   LIGHT_BARRIER_17_STATUS := FALSE;
   LIGHT_BARRIER_18_STATUS := FALSE;
   LIGHT_BARRIER_19_STATUS := FALSE;
   LIGHT_BARRIER_20_STATUS := FALSE;
   LIGHT_BARRIER_21_STATUS := FALSE;
   LIGHT_BARRIER_22_STATUS := FALSE;
   LIGHT_BARRIER_23_STATUS := FALSE;
   LIGHT_BARRIER_24_STATUS := FALSE;
   LIGHT_BARRIER_25_STATUS := FALSE;
   LIGHT_BARRIER_26_STATUS := FALSE;
   LIGHT_BARRIER_27_STATUS := FALSE;
   LIGHT_BARRIER_28_STATUS := FALSE;
   LIGHT_BARRIER_29_STATUS := FALSE;
   LIGHT_BARRIER_30_STATUS := FALSE;
   LIGHT_BARRIER_31_STATUS := FALSE;
   LIGHT_BARRIER_32_STATUS := FALSE;
   PROX_9_STATUS := FALSE;
   PROX_10_STATUS := FALSE;
   PROX_11_STATUS := FALSE;
   PROX_12_STATUS := FALSE;
   PROX_13_STATUS := FALSE;
   PROX_14_STATUS := FALSE;
   PROX_15_STATUS := FALSE;
   PROX_16_STATUS := FALSE;
   PROX_17_STATUS := FALSE;
   PROX_18_STATUS := FALSE;
   PROX_19_STATUS := FALSE;
   PROX_20_STATUS := FALSE;
   PROX_21_STATUS := FALSE;
   PROX_22_STATUS := FALSE;
   PROX_23_STATUS := FALSE;
   PROX_24_STATUS := FALSE;
   FP131 := FALSE;
   FP132 := FALSE;
   FP133 := FALSE;
   FP134 := FALSE;
   FP135 := FALSE;
   TURNTABLE_DELIV_POSITION := FALSE;
   TURNTABLE_REVERSE_ARROW := FALSE;
   TURNTABLE_DIR_SELECT_SW := FALSE;
   TURNTABLE_FLICK_MOTION := FALSE;
   FP140 := FALSE;
   FP141 := FALSE;
   FP142 := FALSE;
   FP143 := FALSE;
   PROX_1_STATUS := FALSE;
   PROX_2_STATUS := FALSE;
   PROX_3_STATUS := FALSE;
   PROX_4_STATUS := FALSE;
   PROX_5_STATUS := FALSE;
   PROX_6_STATUS := FALSE;
   PROX_7_STATUS := FALSE;
   PROX_8_STATUS := FALSE;
   BIT152 := FALSE;
   BIT153 := FALSE;
   BIT154 := FALSE;
   BIT155 := FALSE;
   BIT156 := FALSE;
   BIT157 := FALSE;
   BIT158 := FALSE;
   BIT159 := FALSE;
   SERVICE_SSW_MAIN := FALSE;
   SERVICE_SSW_STATUS := FALSE;
   CLEARING_SSW_MAIN := FALSE;
   CLEARING_SSW_STATUS := FALSE;
   MAN_FEED_SSW_MAIN := FALSE;
   MAN_FEED_SSW_STATUS := FALSE;
   TURNTABLE_SSW_MAIN := FALSE;
   TURNTABLE_SSW_STATUS := FALSE;
   FLIPPER_SSW_MAIN := FALSE;
   FLIPPER_SSW_STATUS := FALSE;
   ROLLER_SSW_MAIN := FALSE;
   ROLLER_SSW_STATUS := FALSE;
   ELEVATOR_ROUND_TRIP_SSW := FALSE;
   BIT173 := FALSE;
   BIT174 := FALSE;
   BIT175 := FALSE;
   HMI_PUSHER_0_TEST_SSW := FALSE;
   HMI_ELEVATOR_SERVICE_SSW := FALSE;
   HMI_ELEVATOR_TEST_DN_SSW := FALSE;
   HMI_ELEVATOR_TEST_UP_SSW := FALSE;
   HMI_ROLLER_TEST_FWD_SSW := FALSE;
   HMI_ROLLER_TEST_REV_SSW := FALSE;
   HMI_PUSHER_1_TEST_SSW := FALSE;
   HMI_CONVEYOR_1_TEST_SSW := FALSE;
   HMI_CONVEYOR_2B_TEST_SSW := FALSE;
   HMI_CONVEYOR_2L_TEST_SSW := FALSE;
   HMI_CONVEYOR_2R_TEST_SSW := FALSE;
   HMI_CONVEYOR_3_TEST_SSW := FALSE;
   HMI_CONVEYOR_4_TEST_SSW := FALSE;
   HMI_CONVEYOR_5_TEST_SSW := FALSE;
   HMI_CONVEYOR_6_TEST_SSW := FALSE;
   HMI_CONVEYOR_7_TEST_SSW := FALSE;
   HMI_CONVEYOR_8_TEST_SSW := FALSE;
   HMI_TURNTABLE_CCW_SSW := FALSE;
   HMI_TURNTABLE_CW_SSW := FALSE;
   HMI_FLIPPER_SERVICE_SSW := FALSE;
   HMI_FLIPPER_FLIP_SSW := FALSE;
   HMI_CONVEYOR_9_TEST_SSW := FALSE;
   HMI_PUSHER_2_TEST_SSW := FALSE;
   HMI_PIVOT_SERVICE_SSW := FALSE;
   HMI_PIVOT_TEST_DN_SSW := FALSE;
   HMI_PIVOT_TEST_UP_SSW := FALSE;
   BIT202 := FALSE;
   BIT203 := FALSE;
   TURNTABLE_SERVICE_PBSHOW := FALSE;
   TURNTABLE_SERVICE_SSW := FALSE;
   HMI_CONVEYOR_10_TEST_SSW := FALSE;
   LOADER_FING_SERVICE_SSW := FALSE;
   LOADER_LIFT_SERVICE_SSW := FALSE;
   LOADER_LIFT_TOP_PB := FALSE;
   LOADER_LIFT_UP_PB := FALSE;
   LOADER_LIFT_DN_PB := FALSE;
   FINGER_RETRACT_TEST_PB := FALSE;
   FINGER_EXTEND_TEST_PB := FALSE;
   FINGER_TILT_TEST_PB := FALSE;
   FINGER_BELT_TEST_SW := FALSE;
   HMI_CONVEYOR_11_TEST_SSW := FALSE;
   HMI_CONVEYOR_12_TEST_SSW := FALSE;
   HMI_CONVEYOR_13_TEST_SSW := FALSE;
   HMI_CONVEYOR_21_TEST_SSW := FALSE;
   HMI_CONVEYOR_22_TEST_SSW := FALSE;
   HMI_CONVEYOR_23_TEST_SSW := FALSE;
   CONVEYOR_0_MOTOR_STATUS := FALSE;
   PUSHER_0_MOTOR_STATUS := FALSE;
   PUSHER_0_COLOR_WORD := W#16#0;
   CONV_0_COLOR_WORD := W#16#0;
   ELEVATOR_COLOR_WORD := W#16#3226;
   PUSHER_1_COLOR_WORD := W#16#0;
   CONV_1_COLOR_WORD := W#16#0;
   CONV_2_BELT_COLOR_WORD := W#16#0;
   LIFT_ROLLER_2_COLOR_WORD := W#16#0;
   CONV_2_ROLLER_COLOR_WORD := W#16#0;
   CONV_3_COLOR_WORD := W#16#0;
   CONV_4_COLOR_WORD := W#16#0;
   CONV_5_COLOR_WORD := W#16#0;
   CONV_6_COLOR_WORD := W#16#0;
   CONV_7_COLOR_WORD := W#16#0;
   FLIPPER_COLOR_WORD := W#16#0;
   CONV_8_COLOR_WORD := W#16#0;
   TURN_TABLE_COLOR_WORD := W#16#0;
   CONV_9_COLOR_WORD := W#16#0;
   PUSHER_2_COLOR_WORD := W#16#0;
   CONV_10_COLOR_WORD := W#16#0;
   CONV_11_COLOR_WORD := W#16#0;
   CONV_12_COLOR_WORD := W#16#0;
   CONV_13_COLOR_WORD := W#16#0;
   CONV_21_COLOR_WORD := W#16#0;
   CONV_22_COLOR_WORD := W#16#0;
   CONV_23_COLOR_WORD := W#16#0;
   LOADER_LIFT_COLOR_WORD := W#16#0;
   LOADER_FING_COLOR_WORD := W#16#0;
   FINGERS_BELT_COLOR_WORD := W#16#0;
   HIGH_LEVEL_23_GRAPHIC := W#16#0;
   LOW_LEVEL_13_GRAPHIC := W#16#0;
   PIVOT_GRAPHIC := W#16#0;
   CONV_3_COUNT := W#16#6;
   CONV_4_COUNT := W#16#0;
   CONV_5_COUNT := W#16#0;
   CONV_6_COUNT := W#16#0;
   CONV_10_COUNT := W#16#0;
   CONV_11_COUNT := W#16#0;
   CONV_12_COUNT := W#16#0;
   CONV_13_COUNT := W#16#0;
   CONV_21_COUNT := W#16#0;
   CONV_22_COUNT := W#16#0;
   CONV_23_COUNT := W#16#0;
   FLIPPER_CCW := W#16#0;
   FLIPPER_CW := W#16#0;
   FLIPPER_POSITION := W#16#0;
   TURN_COLOR := W#16#0;
   FLIPPER_COLOR := W#16#0;
   FLIPPER_PACK_PRESENCE := W#16#0;
   TURNTABLE_PACK_PRESENCE := W#16#0;
   ROLLER_PACK_PRESENCE := W#16#0;
   PUSHER_PACK_PRESENCE := W#16#0;
   CONV_0_STATUS := FALSE;
   PUSHER_0_STATUS := FALSE;
   ELEVATOR_STATUS := FALSE;
   PUSHER_1_STATUS := FALSE;
   CONV_1_STATUS := FALSE;
   TURNTABLE_RNDTRIP := FALSE;
   RNDTRIP_PB_VISIBLE := FALSE;
   BOOL_SPARE227 := FALSE;
   SCREEN_CALL_0 := FALSE;
   SCREEN_CALL_1 := FALSE;
   SCREEN_CALL_2 := FALSE;
   SCREEN_CALL_3 := FALSE;
   SCREEN_CALL_4 := FALSE;
   BOOL_SPARE2276 := FALSE;
   BOOL_SPARE2277 := FALSE;
   BOOL_SPARE2278 := FALSE;
   BOOL_SPARE2279 := FALSE;
   BOOL_SPARE22710 := FALSE;
   BOOL_SPARE22711 := FALSE;
   BOOL_SPARE22712 := FALSE;
   BOOL_SPARE22713 := FALSE;
   BOOL_SPARE22714 := FALSE;
   BOOL_SPARE22715 := FALSE;
   BOOL_SPARE22716 := FALSE;
   BOOL_SPARE22717 := FALSE;
   BOOL_SPARE22718 := FALSE;
   BOOL_SPARE22719 := FALSE;
   BOOL_SPARE22720 := FALSE;
   BOOL_SPARE22721 := FALSE;
   BOOL_SPARE22722 := FALSE;
   BOOL_SPARE22723 := FALSE;
   BOOL_SPARE22724 := FALSE;
   WORD_SPARE23 := W#16#0;
   FLIPPER_TURN_COLOR := W#16#0;
   NEW_ORDER_COLOR := W#16#0;
   SERVICE_FLIPPER := FALSE;
   FLIP_TEST := FALSE;
   SERVICE_TURNTABLE := FALSE;
   TURN_TEST_CW := FALSE;
   TURN_TEST_CCW := FALSE;
   PUSHER_2_TEST := FALSE;
   CONVEYOR_10_TEST_SW := FALSE;
   PIVOT_SERVICE_SW := FALSE;
   PIVOT_UP_TEST_PB := FALSE;
   PIVOT_DN_TEST_PB := FALSE;
   PIVOT_STATUS := FALSE;
   CONV_8_INVERT_SELECT := FALSE;
   CONVEYOR_11_TEST_SW := FALSE;
   CONVEYOR_12_TEST_SW := FALSE;
   CONVEYOR_13_TEST_SW := FALSE;
   CONVEYOR_21_TEST_SW := FALSE;
   CONVEYOR_22_TEST_SW := FALSE;
   CONVEYOR_23_TEST_SW := FALSE;
   LOADER_SERVICE_SW := FALSE;
   LOADER_UP_TEST_PB := FALSE;
   LOADER_DN_TEST_PB := FALSE;
   FINGERS_EXTEND_TEST_PB := FALSE;
   FINGERS_RETRACT_TEST_PB := FALSE;
   FP_ONESHOT_0 := FALSE;
   CONVEYOR_0_SERVICE_SW := FALSE;
   ELEVATOR_SERVICE_SW := FALSE;
   CONVEYOR_1_SERVICE_SW := FALSE;
   CONVEYOR_2_SERVICE_SW := FALSE;
   CONVEYOR_3_SERVICE_SW := FALSE;
   CONVEYOR_4_SERVICE_SW := FALSE;
   CONVEYOR_5_SERVICE_SW := FALSE;
   CONVEYOR_6_SERVICE_SW := FALSE;
   CONVEYOR_7_SERVICE_SW := FALSE;
   CONVEYOR_8_SERVICE_SW := FALSE;
   CONVEYOR_9_SERVICE_SW := FALSE;
   CONVEYOR_10_SERVICE_SW := FALSE;
   CONVEYOR_11_SERVICE_SW := FALSE;
   CONVEYOR_21_SERVICE_SW := FALSE;
   LOADER_SERVICE_ENABLE_SW := FALSE;
   CTRL48 := FALSE;
   CTRL49 := FALSE;
   CTRL50 := FALSE;
   CTRL51 := FALSE;
   CTRL52 := FALSE;
   CTRL53 := FALSE;
   CTRL54 := FALSE;
   CTRL55 := FALSE;
   CTRL56 := FALSE;
   CLEARING_FUNCTION := W#16#0;
   WORD57 := W#16#0;
   WORD58 := W#16#0;
   ACTUAL_HMI_SCREEN_NO := W#16#0;
   CONVEYOR_MAXCOUNT_L := W#16#6;
   CONVEYOR_MAXCOUNT_W := W#16#7;
   WORD62 := W#16#0;
   CONV_7_POS_mS := W#16#96;
   CONV_8_POS_FWD_mS := W#16#0;
   CONV_8_POS_REV_mS := W#16#0;
   CONV_9_POS_mS := W#16#0;
   WORD_PACKET_LENGTH := W#16#0;
   DELAY_DISPLAY_7 := W#16#0;
   DELAY_DISPLAY_9 := W#16#0;
   WORD_SPARE2 := W#16#0;
   WORD_SPARE3 := W#16#0;
   WORD_SPARE4 := W#16#0;
END_DATA_BLOCK

DATA_BLOCK "DB LAUER"
TITLE =
VERSION : 0.0


  STRUCT
   D_0 : WORD ;
   D_1 : WORD ;
   D_2 : WORD ;
   D_3 : WORD  := W#16#A1;
   D_4 : WORD ;
   D_5 : WORD ;
   D_6 : WORD ;
   D_7 : WORD ;
   D_8 : WORD ;
   D_9 : WORD  := W#16#2006;
   D_10 : WORD  := W#16#1023;
   D_11 : WORD  := W#16#13;
   D_12 : WORD  := W#16#3439;
   D_13 : WORD  := W#16#3500;
   D_14 : WORD ;
   D_15 : WORD  := W#16#1A0;
   D_16 : WORD ;
   D_17 : WORD ;
   D_18 : WORD  := W#16#7C02;
   D_19 : WORD ;
   D_20 : WORD ;
   D_21 : WORD ;
   D_22 : WORD ;
   D_23 : WORD ;
   D_24 : WORD  := W#16#8480;
   D_25 : WORD ;
   D_26 : WORD ;
   D_27 : WORD ;
   D_28 : WORD ;
   D_29 : WORD ;
   D_30 : WORD ;
   D_31 : WORD ;
   D_32 : WORD ;
   D_33 : WORD ;
   D_34 : WORD ;
   D_35 : WORD ;
   D_36 : WORD  := W#16#F00;
   D_37 : WORD  := W#16#3001;
   D_38 : WORD ;
   D_39 : WORD ;
   D_40 : WORD ;
   D_41 : WORD ;
   D_42 : WORD ;
   D_43 : WORD ;
   D_44 : WORD ;
   D_45 : WORD ;
   D_46 : WORD ;
   D_47 : WORD ;
   D_48 : WORD ;
   D_49 : WORD ;
   D_50 : WORD ;
   D_51 : WORD ;
   D_52 : WORD ;
   D_53 : WORD ;
   D_54 : WORD ;
   D_55 : WORD ;
   D_56 : WORD ;
   D_57 : WORD ;
   D_58 : WORD ;
   D_59 : WORD ;
   D_60 : WORD ;
   D_61 : WORD ;
   D_62 : WORD ;
   D_63 : WORD ;
   D_64 : WORD ;
   D_65 : WORD ;
   D_66 : WORD ;
   D_67 : WORD ;
   D_68 : WORD ;
   D_69 : WORD ;
   D_70 : WORD ;
   D_71 : WORD ;
   D_72 : WORD ;
   D_73 : WORD ;
   D_74 : WORD ;
   D_75 : WORD ;
   D_76 : WORD ;
   D_77 : WORD  := W#16#4;
   D_78 : WORD  := W#16#2;
   D_79 : WORD  := W#16#1;
   D_80 : WORD  := W#16#1;
   D_81 : WORD  := W#16#1;
   D_82 : WORD  := W#16#1;
   D_83 : WORD  := W#16#1;
   D_84 : WORD  := W#16#2;
   D_85 : WORD  := W#16#3;
   D_86 : WORD  := W#16#2;
   D_87 : WORD  := W#16#1;
   D_88 : WORD  := W#16#1;
   D_89 : WORD  := W#16#3;
   D_90 : WORD  := W#16#4;
   D_91 : WORD  := W#16#7;
   D_92 : WORD  := W#16#9;
   D_93 : WORD  := W#16#3;
   D_94 : WORD  := W#16#3;
   D_95 : WORD  := W#16#4;
   D_96 : WORD  := W#16#1;
   D_97 : WORD  := W#16#1;
   D_98 : WORD  := W#16#1;
   D_99 : WORD  := W#16#1;
   D_100 : WORD  := W#16#1;
   D_101 : WORD  := W#16#1;
   D_102 : WORD  := W#16#1;
   D_103 : WORD ;
   D_104 : WORD ;
   D_105 : WORD ;
   D_106 : WORD ;
   D_107 : WORD ;
   D_108 : WORD ;
   D_109 : WORD ;
   D_110 : WORD  := W#16#2;
   D_111 : WORD ;
   D_112 : WORD ;
   D_113 : WORD ;
   D_114 : WORD ;
   D_115 : WORD ;
   D_116 : WORD ;
   D_117 : WORD  := W#16#7;
   D_118 : WORD  := W#16#1;
   D_119 : WORD  := W#16#1;
   D_120 : WORD  := W#16#2010;
   D_121 : WORD  := W#16#58;
   D_122 : WORD  := W#16#2010;
   D_123 : WORD  := W#16#2090;
   D_124 : WORD  := W#16#9;
   D_125 : WORD ;
   D_126 : WORD  := W#16#15;
   D_127 : WORD ;
   D_128 : WORD ;
   D_129 : WORD  := W#16#6;
   D_130 : WORD  := W#16#320;
   D_131 : WORD ;
   D_132 : WORD  := W#16#B7;
   D_133 : WORD  := W#16#1EDE;
   D_134 : WORD ;
   D_135 : WORD ;
   D_136 : WORD ;
   D_137 : WORD ;
   D_138 : WORD ;
   D_139 : WORD ;
   D_140 : WORD  := W#16#320;
   D_141 : WORD ;
   D_142 : WORD  := W#16#37;
   D_143 : WORD  := W#16#5D2;
   D_144 : WORD ;
   D_145 : WORD ;
   D_146 : WORD ;
   D_147 : WORD ;
   D_148 : WORD ;
   D_149 : WORD ;
   D_150 : WORD  := W#16#5C;
   D_151 : WORD ;
   D_152 : WORD ;
   D_153 : WORD ;
   D_154 : WORD ;
   D_155 : WORD ;
   D_156 : WORD ;
   D_157 : WORD ;
   D_158 : WORD ;
   D_159 : WORD ;
   D_160 : WORD  := W#16#320;
   D_161 : WORD ;
   D_162 : WORD  := W#16#B9;
   D_163 : WORD  := W#16#181F;
   D_164 : WORD ;
   D_165 : WORD ;
   D_166 : WORD ;
   D_167 : WORD ;
   D_168 : WORD ;
   D_169 : WORD ;
   D_170 : WORD  := W#16#320;
   D_171 : WORD ;
   D_172 : WORD  := W#16#F;
   D_173 : WORD  := W#16#14B9;
   D_174 : WORD ;
   D_175 : WORD ;
   D_176 : WORD ;
   D_177 : WORD ;
   D_178 : WORD ;
   D_179 : WORD ;
   D_180 : WORD  := W#16#320;
   D_181 : WORD ;
   D_182 : WORD ;
   D_183 : WORD  := W#16#4B0;
   D_184 : WORD  := W#16#1;
   D_185 : WORD  := W#16#1;
   D_186 : WORD ;
   D_187 : WORD ;
   D_188 : WORD ;
   D_189 : WORD ;
   D_190 : WORD ;
   D_191 : WORD ;
   D_192 : WORD ;
   D_193 : WORD ;
   D_194 : WORD ;
   D_195 : WORD ;
   D_196 : WORD ;
   D_197 : WORD ;
   D_198 : WORD ;
   D_199 : WORD ;
   D_200 : WORD ;
   D_201 : WORD ;
   D_202 : WORD ;
   D_203 : WORD ;
   D_204 : WORD ;
   D_205 : WORD ;
   D_206 : WORD ;
   D_207 : WORD ;
   D_208 : WORD ;
   D_209 : WORD ;
   D_210 : WORD ;
   D_211 : WORD ;
   D_212 : WORD ;
   D_213 : WORD ;
   D_214 : WORD ;
   D_215 : WORD ;
   D_216 : WORD ;
   D_217 : WORD ;
   D_218 : WORD ;
   D_219 : WORD ;
   D_220 : WORD ;
   D_221 : WORD ;
   D_222 : WORD ;
   D_223 : WORD ;
   D_224 : WORD ;
   D_225 : WORD ;
   D_226 : WORD ;
   D_227 : WORD ;
   D_228 : WORD ;
   D_229 : WORD ;
   D_230 : WORD ;
   D_231 : WORD ;
   D_232 : WORD ;
   D_233 : WORD ;
   D_234 : WORD ;
   D_235 : WORD ;
   D_236 : WORD ;
   D_237 : WORD ;
   D_238 : WORD ;
   D_239 : WORD ;
   D_240 : WORD ;
   D_241 : WORD ;
   D_242 : WORD ;
   D_243 : WORD ;
   D_244 : WORD ;
   D_245 : WORD ;
   D_246 : WORD ;
   D_247 : WORD ;
   D_248 : WORD ;
   D_249 : WORD ;
   D_250 : WORD ;
   D_251 : WORD ;
   D_252 : WORD  := W#16#58;
   D_253 : WORD  := W#16#9;
   D_254 : WORD ;
   D_255 : WORD  := W#16#12;
  END_STRUCT ;
BEGIN
   D_0 := W#16#4B;
   D_1 := W#16#0;
   D_2 := W#16#0;
   D_3 := W#16#0;
   D_4 := W#16#0;
   D_5 := W#16#0;
   D_6 := W#16#0;
   D_7 := W#16#0;
   D_8 := W#16#0;
   D_9 := W#16#2010;
   D_10 := W#16#527;
   D_11 := W#16#619;
   D_12 := W#16#306;
   D_13 := W#16#3F00;
   D_14 := W#16#0;
   D_15 := W#16#1A0;
   D_16 := W#16#0;
   D_17 := W#16#0;
   D_18 := W#16#7C02;
   D_19 := W#16#0;
   D_20 := W#16#0;
   D_21 := W#16#0;
   D_22 := W#16#0;
   D_23 := W#16#0;
   D_24 := W#16#8480;
   D_25 := W#16#0;
   D_26 := W#16#0;
   D_27 := W#16#0;
   D_28 := W#16#0;
   D_29 := W#16#0;
   D_30 := W#16#0;
   D_31 := W#16#0;
   D_32 := W#16#0;
   D_33 := W#16#0;
   D_34 := W#16#0;
   D_35 := W#16#0;
   D_36 := W#16#F00;
   D_37 := W#16#3001;
   D_38 := W#16#0;
   D_39 := W#16#0;
   D_40 := W#16#0;
   D_41 := W#16#0;
   D_42 := W#16#0;
   D_43 := W#16#0;
   D_44 := W#16#0;
   D_45 := W#16#0;
   D_46 := W#16#0;
   D_47 := W#16#0;
   D_48 := W#16#0;
   D_49 := W#16#0;
   D_50 := W#16#0;
   D_51 := W#16#0;
   D_52 := W#16#0;
   D_53 := W#16#0;
   D_54 := W#16#0;
   D_55 := W#16#0;
   D_56 := W#16#0;
   D_57 := W#16#0;
   D_58 := W#16#0;
   D_59 := W#16#0;
   D_60 := W#16#0;
   D_61 := W#16#0;
   D_62 := W#16#0;
   D_63 := W#16#0;
   D_64 := W#16#0;
   D_65 := W#16#0;
   D_66 := W#16#0;
   D_67 := W#16#0;
   D_68 := W#16#0;
   D_69 := W#16#0;
   D_70 := W#16#0;
   D_71 := W#16#0;
   D_72 := W#16#0;
   D_73 := W#16#0;
   D_74 := W#16#0;
   D_75 := W#16#0;
   D_76 := W#16#0;
   D_77 := W#16#4;
   D_78 := W#16#2;
   D_79 := W#16#4;
   D_80 := W#16#1;
   D_81 := W#16#1;
   D_82 := W#16#1;
   D_83 := W#16#1;
   D_84 := W#16#A;
   D_85 := W#16#4;
   D_86 := W#16#9;
   D_87 := W#16#1;
   D_88 := W#16#1;
   D_89 := W#16#1;
   D_90 := W#16#4;
   D_91 := W#16#7;
   D_92 := W#16#9;
   D_93 := W#16#4;
   D_94 := W#16#2;
   D_95 := W#16#1;
   D_96 := W#16#0;
   D_97 := W#16#0;
   D_98 := W#16#0;
   D_99 := W#16#0;
   D_100 := W#16#0;
   D_101 := W#16#1;
   D_102 := W#16#0;
   D_103 := W#16#0;
   D_104 := W#16#0;
   D_105 := W#16#0;
   D_106 := W#16#0;
   D_107 := W#16#0;
   D_108 := W#16#0;
   D_109 := W#16#0;
   D_110 := W#16#2;
   D_111 := W#16#0;
   D_112 := W#16#0;
   D_113 := W#16#0;
   D_114 := W#16#C;
   D_115 := W#16#C;
   D_116 := W#16#1;
   D_117 := W#16#7;
   D_118 := W#16#0;
   D_119 := W#16#1;
   D_120 := W#16#2010;
   D_121 := W#16#96;
   D_122 := W#16#2010;
   D_123 := W#16#2090;
   D_124 := W#16#C;
   D_125 := W#16#0;
   D_126 := W#16#15;
   D_127 := W#16#0;
   D_128 := W#16#0;
   D_129 := W#16#6;
   D_130 := W#16#320;
   D_131 := W#16#0;
   D_132 := W#16#2A9;
   D_133 := W#16#238;
   D_134 := W#16#0;
   D_135 := W#16#0;
   D_136 := W#16#0;
   D_137 := W#16#0;
   D_138 := W#16#0;
   D_139 := W#16#0;
   D_140 := W#16#320;
   D_141 := W#16#0;
   D_142 := W#16#98;
   D_143 := W#16#1262;
   D_144 := W#16#0;
   D_145 := W#16#0;
   D_146 := W#16#0;
   D_147 := W#16#0;
   D_148 := W#16#0;
   D_149 := W#16#0;
   D_150 := W#16#67;
   D_151 := W#16#0;
   D_152 := W#16#0;
   D_153 := W#16#0;
   D_154 := W#16#0;
   D_155 := W#16#0;
   D_156 := W#16#0;
   D_157 := W#16#0;
   D_158 := W#16#0;
   D_159 := W#16#0;
   D_160 := W#16#320;
   D_161 := W#16#0;
   D_162 := W#16#2C1;
   D_163 := W#16#FD0;
   D_164 := W#16#0;
   D_165 := W#16#0;
   D_166 := W#16#0;
   D_167 := W#16#0;
   D_168 := W#16#0;
   D_169 := W#16#0;
   D_170 := W#16#320;
   D_171 := W#16#0;
   D_172 := W#16#0;
   D_173 := W#16#0;
   D_174 := W#16#1;
   D_175 := W#16#1;
   D_176 := W#16#0;
   D_177 := W#16#0;
   D_178 := W#16#0;
   D_179 := W#16#0;
   D_180 := W#16#320;
   D_181 := W#16#0;
   D_182 := W#16#0;
   D_183 := W#16#7B0;
   D_184 := W#16#1;
   D_185 := W#16#1;
   D_186 := W#16#0;
   D_187 := W#16#0;
   D_188 := W#16#0;
   D_189 := W#16#0;
   D_190 := W#16#0;
   D_191 := W#16#0;
   D_192 := W#16#0;
   D_193 := W#16#0;
   D_194 := W#16#0;
   D_195 := W#16#0;
   D_196 := W#16#0;
   D_197 := W#16#0;
   D_198 := W#16#0;
   D_199 := W#16#0;
   D_200 := W#16#0;
   D_201 := W#16#0;
   D_202 := W#16#0;
   D_203 := W#16#0;
   D_204 := W#16#0;
   D_205 := W#16#0;
   D_206 := W#16#0;
   D_207 := W#16#0;
   D_208 := W#16#0;
   D_209 := W#16#0;
   D_210 := W#16#0;
   D_211 := W#16#0;
   D_212 := W#16#0;
   D_213 := W#16#0;
   D_214 := W#16#0;
   D_215 := W#16#0;
   D_216 := W#16#0;
   D_217 := W#16#0;
   D_218 := W#16#0;
   D_219 := W#16#0;
   D_220 := W#16#0;
   D_221 := W#16#0;
   D_222 := W#16#0;
   D_223 := W#16#0;
   D_224 := W#16#0;
   D_225 := W#16#0;
   D_226 := W#16#0;
   D_227 := W#16#0;
   D_228 := W#16#0;
   D_229 := W#16#0;
   D_230 := W#16#0;
   D_231 := W#16#0;
   D_232 := W#16#0;
   D_233 := W#16#0;
   D_234 := W#16#0;
   D_235 := W#16#0;
   D_236 := W#16#0;
   D_237 := W#16#0;
   D_238 := W#16#0;
   D_239 := W#16#0;
   D_240 := W#16#0;
   D_241 := W#16#0;
   D_242 := W#16#0;
   D_243 := W#16#0;
   D_244 := W#16#0;
   D_245 := W#16#0;
   D_246 := W#16#0;
   D_247 := W#16#0;
   D_248 := W#16#0;
   D_249 := W#16#0;
   D_250 := W#16#0;
   D_251 := W#16#0;
   D_252 := W#16#C;
   D_253 := W#16#12;
   D_254 := W#16#0;
   D_255 := W#16#12;
END_DATA_BLOCK

FUNCTION "LAUER TIME" : VOID
TITLE =
// TIMER
NAME : _TIMER
VERSION : 0.0


VAR_OUTPUT
  QUEL : WORD ;	// QUEL
  _TIME : WORD ;	// TIME
END_VAR
BEGIN
NETWORK
TITLE =

      OPN   "DB LAUER";
      L     #QUEL;
      T     DBW  504;

      L     DBW  504;
      ITB   ;
      T     DBW  506;

      L     DBW  506;
      T     #_TIME;
END_FUNCTION

FUNCTION "SENSOR CHECK" : VOID
TITLE =Sensor Check
//Counting Foul Sensor Switching of less than PreSet Time (500mS)
VERSION : 0.1


VAR_INPUT
  Bit : BOOL ;
  Preset_ms : INT ;
  Plc_Scan_ms : INT ;
END_VAR
VAR_IN_OUT
  Rising_Pulse_1 : BOOL ;	//Db3 Struct
  Rising_Pulse_2 : BOOL ;	//Db3 Struct
  Memory_Bit_1 : BOOL ;	//Db3 Struct
  Memory_Bit_2 : BOOL ;	//Db3 Struct
  Word_Buffer : INT ;	//Db3 Struct
  Word_Result : INT ;	//Db3 Struct
END_VAR
VAR_TEMP
  MEMORY_BIT : BOOL ;
  Bool2 : BOOL ;
  Bool3 : BOOL ;
  Bool4 : BOOL ;
  Bool5 : BOOL ;
  Bool6 : BOOL ;
  Bool7 : BOOL ;
  Bool8 : BOOL ;
END_VAR
BEGIN
NETWORK
TITLE =Input Bit - Reset
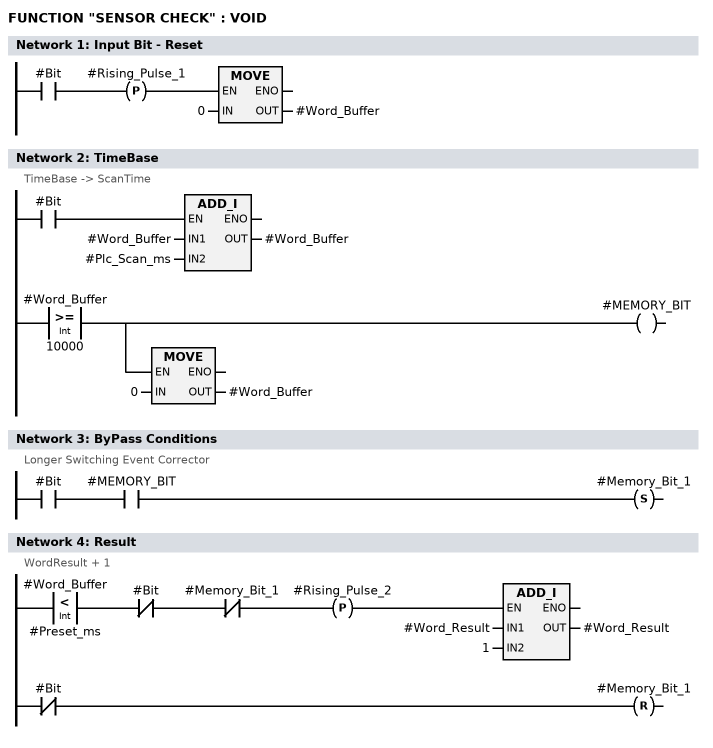

      A     #Bit;
      FP    #Rising_Pulse_1;
      JNB   _001;
      L     0;
      T     #Word_Buffer;

_001: NOP   0;
NETWORK
TITLE =TimeBase
//TimeBase -> ScanTime
      A     #Bit;
      JNB   _002;
      L     #Word_Buffer;
      L     #Plc_Scan_ms;
      +I    ;
      T     #Word_Buffer;

_002: NOP   0;

      A(    ;
      L     #Word_Buffer;
      L     10000;
      >=I   ;
      )     ;
      =     #MEMORY_BIT;
      JNB   _003;
      L     0;
      T     #Word_Buffer;

_003: NOP   0;
NETWORK
TITLE =ByPass Conditions
//Longer Switching Event Corrector

      A     #Bit;
      A     #MEMORY_BIT;
      S     #Memory_Bit_1;
NETWORK
TITLE =Result
//WordResult + 1
      A(    ;
      L     #Word_Buffer;
      L     #Preset_ms;
      <I    ;
      )     ;
      AN    #Bit;
      AN    #Memory_Bit_1;
      FP    #Rising_Pulse_2;
      JNB   _004;
      L     #Word_Result;
      L     1;
      +I    ;
      T     #Word_Result;

_004: NOP   0;

      AN    #Bit;
      R     #Memory_Bit_1;

END_FUNCTION

FUNCTION "DE-BOUNCER / COUNTER" : VOID
TITLE =Packet De-Bouncer / Counter  FC8
//==========================================================================
//  PACKET DE-BOUNCER / COUNTER  -  v0.7  (Replaces FC6 "DE-BOUNCER OLD")
//
//  COUNT UP   (Bit_0 = InFeed Sensor, gated by the caller)
//    - Bit_0 ON time is added while the packet is under the sensor.
//    - +1 once the ON time reaches Preset_MIN_mS.
//    - Re-armed only after Bit_0 stays OFF for the Gap time, so a
//      "U" shaped packet (short opening) is counted ONCE.
//    - A blip shorter than Preset_MIN_mS is dropped at the Gap.
//
//  COUNT DOWN (Bit_1 = RAW Exit Sensor, Transfer_Start = Transfer Step)
//    - Bit_1 ON time is only added while Transfer_Start is ON
//      (a packet parked on the exit sensor is NOT counted).
//    - -1 when the packet has LEFT: Bit_1 OFF for the Gap time and
//      ON time >= Preset_MIN_mS.
//    - Butted packets (exit sensor never clears): -1 every
//      HighSpd_Dimension_mS + Gap of continuous ON time.
//      HighSpd_Dimension_mS = 0 disables this.
//
//  Gap = Space_DX_mS / 2  (min 100 mS)
//
//  HMI (Word_Count, In/Out)
//    - Operator edit or external reset (write 0) is taken over on the
//      next call, as FC6 did.  Result is written back every call.
//
//  ERROR
//    - Bit_0 continuously ON >= 5 s -> IO_DB.Error / Q_Error (latched).
//    - Cleared by Error_Reset.
//
//  Call while the conveyor runs + ~1 s off-delay.
//  ReSample_DX, Conveyor_Type, LowSpd_Dimension_mS: kept for interface
//  compatibility, not used.
//==========================================================================
VERSION : 0.7


VAR_INPUT
  Bit_0 : BOOL ;	//InFeed Sensor - Count UP (gated by caller)
  Bit_1 : BOOL ;	//Exit Sensor - Count DOWN (RAW sensor)
  Transfer_Start : BOOL ;	//Transfer Step Active - Count DOWN Enable
  Error_Reset : BOOL ;	//Fault Reset PB
  Space_DX_mS : INT ;	//Nominal Space Between Packets [mS] - Gap = 50%
  ReSample_DX : INT ;	//Not Used (Compatibility)
  Conveyor_Type : INT ;	//Info Only: 1 Collator, 2 Delivery, 3 Link
  Preset_MIN_mS : INT ;	//Min ON Time to Accept a Packet [mS]
  LowSpd_Dimension_mS : INT ;	//Not Used (Compatibility)
  HighSpd_Dimension_mS : INT ;	//Packet Dimension @ Transfer Speed [mS] - 0 = Off
  Plc_Scan_mS : INT ;	//PLC ScanTime [mS]
END_VAR
VAR_OUTPUT
  Q_Error : BOOL ;	//Bit_0 Stuck
END_VAR
VAR_IN_OUT
  Word_Count : WORD ;	//HMI Packet Count (Read + Write Back) - WORD as in "HMI_DB"
  IO_DB : "Debouncer Counter Struct";
END_VAR
BEGIN
NETWORK
TITLE =Init on First Call - Take Over HMI Count

      AN    #IO_DB.FirstScan_Done;
      JCN   INIT;
      L     0;
      T     #IO_DB.Bit0_Entry_mS;
      T     #IO_DB.Bit0_OFF_mS;
      T     #IO_DB.Bit0_Stuck_mS;
      T     #IO_DB.Bit1_Exit_mS;
      T     #IO_DB.Bit1_OFF_mS;
      L     #Word_Count;
      T     #IO_DB.Count_Result;
      T     #IO_DB.HMI_Last;
      SET   ;
      R     #IO_DB.Bit0_ON_Latch;
      R     #IO_DB.Bit1_ON_Latch;
      R     #IO_DB.Count_Done_Latch_0;
      R     #IO_DB.Error;
      S     #IO_DB.FirstScan_Done;
INIT: NOP   0;
NETWORK
TITLE =HMI Count Changed Outside (Operator Edit / Reset) - Take Over

      L     #Word_Count;
      L     #IO_DB.HMI_Last;
      <>I   ;
      JCN   H001;
      L     #Word_Count;
      T     #IO_DB.Count_Result;
H001: NOP   0;
NETWORK
TITLE =Windows

      L     #Space_DX_mS;
      L     2;
      /I    ;
      T     #IO_DB.Space_Between; // Gap Confirm [mS]
      L     100;
      <I    ;
      JCN   P001;
      L     100;
      T     #IO_DB.Space_Between; // Min 100 mS
P001: L     #Preset_MIN_mS;
      T     #IO_DB.InFeed_Window_mS; // Info
      L     #HighSpd_Dimension_mS;
      L     #IO_DB.Space_Between;
      +I    ;
      T     #IO_DB.Exit_Window_mS; // Butted Packets Window
NETWORK
TITLE =Count UP - InFeed Sensor Timing

      A     #Bit_0;
      JCN   U001;
      SET   ;
      S     #IO_DB.Bit0_ON_Latch; // Packet Seen
      L     0;
      T     #IO_DB.Bit0_OFF_mS;
      L     #IO_DB.Bit0_Entry_mS;
      L     #Plc_Scan_mS;
      +I    ;
      T     #IO_DB.Bit0_Entry_mS; // ON Time - This Packet
      L     #IO_DB.Bit0_Stuck_mS;
      L     #Plc_Scan_mS;
      +I    ;
      T     #IO_DB.Bit0_Stuck_mS; // Continuous ON Time
      JU    U002;
U001: L     0;
      T     #IO_DB.Bit0_Stuck_mS;
      A     #IO_DB.Bit0_ON_Latch;
      JCN   U002;
      L     #IO_DB.Bit0_OFF_mS;
      L     #Plc_Scan_mS;
      +I    ;
      T     #IO_DB.Bit0_OFF_mS; // Gap Time
U002: NOP   0;
NETWORK
TITLE =Count UP - Packet Accepted +1

      A     #IO_DB.Bit0_ON_Latch;
      AN    #IO_DB.Count_Done_Latch_0; // Not Counted Yet
      A(    ;
      L     #IO_DB.Bit0_Entry_mS;
      L     #Preset_MIN_mS;
      >=I   ;
      )     ;
      JCN   U003;
      L     #IO_DB.Count_Result;
      L     1;
      +I    ;
      T     #IO_DB.Count_Result;
      SET   ;
      S     #IO_DB.Count_Done_Latch_0;
U003: NOP   0;
NETWORK
TITLE =Count UP - Gap Confirmed - Re-Arm

      A(    ;
      L     #IO_DB.Bit0_OFF_mS;
      L     #IO_DB.Space_Between;
      >=I   ;
      )     ;
      JCN   U004;
      SET   ;
      R     #IO_DB.Bit0_ON_Latch;
      R     #IO_DB.Count_Done_Latch_0;
      L     0;
      T     #IO_DB.Bit0_Entry_mS;
      T     #IO_DB.Bit0_OFF_mS;
U004: NOP   0;
NETWORK
TITLE =Count DOWN - Exit Sensor Timing

      A     #Bit_1;
      JCN   D001;
      L     0;
      T     #IO_DB.Bit1_OFF_mS;
      A     #Transfer_Start; // ON Time only while Transfering
      JCN   D002;
      SET   ;
      S     #IO_DB.Bit1_ON_Latch;
      L     #IO_DB.Bit1_Exit_mS;
      L     #Plc_Scan_mS;
      +I    ;
      T     #IO_DB.Bit1_Exit_mS; // ON Time - This Packet
      JU    D002;
D001: A     #IO_DB.Bit1_ON_Latch;
      JCN   D002;
      L     #IO_DB.Bit1_OFF_mS;
      L     #Plc_Scan_mS;
      +I    ;
      T     #IO_DB.Bit1_OFF_mS; // Gap Time
D002: NOP   0;
NETWORK
TITLE =Count DOWN - Butted Packets -1 (Exit Sensor Never Clears)
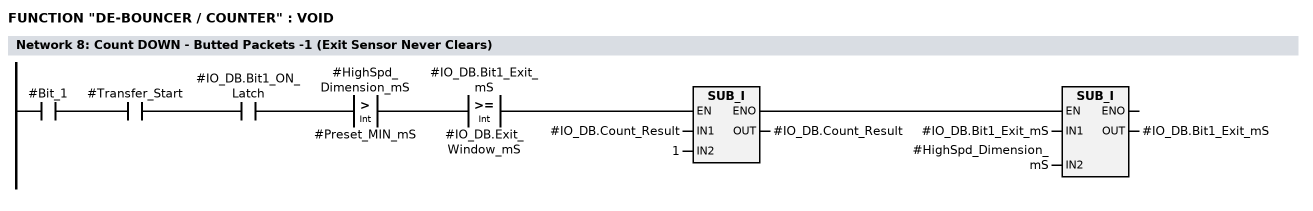

      A     #Bit_1;
      A     #Transfer_Start;
      A     #IO_DB.Bit1_ON_Latch;
      A(    ;
      L     #HighSpd_Dimension_mS;
      L     #Preset_MIN_mS;
      >I    ;
      )     ;
      A(    ;
      L     #IO_DB.Bit1_Exit_mS;
      L     #IO_DB.Exit_Window_mS;
      >=I   ;
      )     ;
      JCN   D003;
      L     #IO_DB.Count_Result;
      L     1;
      -I    ;
      T     #IO_DB.Count_Result;
      L     #IO_DB.Bit1_Exit_mS;
      L     #HighSpd_Dimension_mS;
      -I    ;
      T     #IO_DB.Bit1_Exit_mS; // Keep the Rest for the Next Packet
D003: NOP   0;
NETWORK
TITLE =Count DOWN - Packet Left -1

      A(    ;
      L     #IO_DB.Bit1_OFF_mS;
      L     #IO_DB.Space_Between;
      >=I   ;
      )     ;
      JCN   D005;
      A(    ;
      L     #IO_DB.Bit1_Exit_mS;
      L     #Preset_MIN_mS;
      >=I   ;
      )     ;
      JCN   D004; // Too Short = Not a Packet
      L     #IO_DB.Count_Result;
      L     1;
      -I    ;
      T     #IO_DB.Count_Result;
D004: SET   ;
      R     #IO_DB.Bit1_ON_Latch;
      L     0;
      T     #IO_DB.Bit1_Exit_mS;
      T     #IO_DB.Bit1_OFF_mS;
D005: NOP   0;
NETWORK
TITLE =Timers Overflow Clamp 30s

      L     #IO_DB.Bit0_Entry_mS;
      L     30000;
      >I    ;
      JCN   K001;
      L     30000;
      T     #IO_DB.Bit0_Entry_mS;
K001: L     #IO_DB.Bit0_Stuck_mS;
      L     30000;
      >I    ;
      JCN   K002;
      L     30000;
      T     #IO_DB.Bit0_Stuck_mS;
K002: L     #IO_DB.Bit1_Exit_mS;
      L     30000;
      >I    ;
      JCN   K003;
      L     30000;
      T     #IO_DB.Bit1_Exit_mS;
K003: NOP   0;
NETWORK
TITLE =Clamp Packet Qty  0...Maximum_Count  (Max 0 = No Limit)

      L     #IO_DB.Count_Result;
      L     0;
      <I    ;
      JCN   C001;
      L     0;
      T     #IO_DB.Count_Result;
C001: L     #IO_DB.Maximum_Count;
      L     0;
      >I    ;
      JCN   C002;
      L     #IO_DB.Count_Result;
      L     #IO_DB.Maximum_Count;
      >I    ;
      JCN   C002;
      L     #IO_DB.Maximum_Count;
      T     #IO_DB.Count_Result;
C002: NOP   0;
NETWORK
TITLE =InFeed Sensor Stuck >= 5s - Error
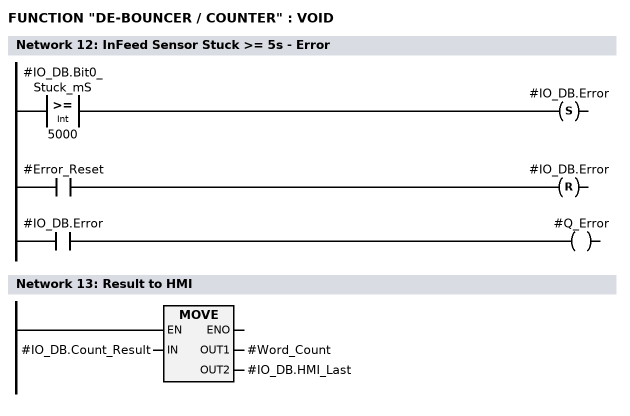

      A(    ;
      L     #IO_DB.Bit0_Stuck_mS;
      L     5000;
      >=I   ;
      )     ;
      S     #IO_DB.Error;
      A     #Error_Reset;
      R     #IO_DB.Error;
      A     #IO_DB.Error;
      =     #Q_Error;
NETWORK
TITLE =Result to HMI

      L     #IO_DB.Count_Result;
      T     #Word_Count;
      T     #IO_DB.HMI_Last;
END_FUNCTION

FUNCTION "SCALER" : REAL
TITLE =Linear interpolation between two points
AUTHOR : APC
FAMILY : CONV_LIB
NAME : LINEAR
VERSION : 1.0


VAR_INPUT
  X : REAL ;	//[-] Input value
  X1 : REAL ;	//[-] First interpolation point, x-value
  Y1 : REAL ;	//[-] First interpolation point, y-value
  X2 : REAL ;	//[-] Second interpolation point, x-value
  Y2 : REAL ;	//[-] Second interpolation point, y-value
END_VAR
VAR_TEMP
  X_CALC_1 : REAL ;	//[-] x1 for Calculation
  Y_CALC_1 : REAL ;	//[-] y1 for Calculation
  X_CALC_2 : REAL ;	//[-] x2 for Calculation
  Y_CALC_2 : REAL ;	//[-] y2 for Calculation
END_VAR
BEGIN
NETWORK
TITLE =SCL network
//compiled by SCL compiler version:  SCLCOMP K05.06.00.00_11.01.00.01 release
//      SET
//     SAVE
//     =     L     16.1
      L     0.000000e+00;
      T     #RET_VAL;
//;
      L     #X1;
      L     #X2;
      <>R   ;
      JCN   A7d0;
//;
      L     #X1;
      L     #X2;
      >R    ;
      JCN   A7d1;
//;
      L     #X2;
      T     #X_CALC_1;
//;
      L     #Y2;
      T     #Y_CALC_1;
//;
      L     #X1;
      T     #X_CALC_2;
//;
      L     #Y1;
      T     #Y_CALC_2;
      JU    A7d2;

A7d1: L     #X1;
      T     #X_CALC_1;
//;
      L     #Y1;
      T     #Y_CALC_1;
//;
      L     #X2;
      T     #X_CALC_2;
//;
      L     #Y2;
      T     #Y_CALC_2;
A7d2: L     #X;

      L     #X_CALC_1;
      <=R   ;
      JCN   A7d3;
      L     #Y_CALC_1;
      T     #RET_VAL;
      JU    A7d0;

A7d3: L     #X;
      L     #X_CALC_2;
      >=R   ;
      JCN   A7d5;
      L     #Y_CALC_2;
      T     #RET_VAL;
      JU    A7d0;

A7d5: L     #X;
      L     #X_CALC_1;
      -R    ;
      L     #X_CALC_2;
      TAK   ;
      T     LD    18;
      TAK   ;
      L     #X_CALC_1;
      -R    ;
      L     LD    18;
      TAK   ;
      /R    ;
      L     #Y_CALC_2;
      TAK   ;
      T     LD    18;
      TAK   ;
      L     #Y_CALC_1;
      -R    ;
      L     LD    18;
      *R    ;
      L     #Y_CALC_1;
      +R    ;
      T     #RET_VAL;

A7d0: CLR   ;

//    A     L     16.1
//    SAVE
//    BE
END_FUNCTION

FUNCTION "LAUER KEYS 1" : VOID
TITLE =
NAME : TASTAUSW
VERSION : 0.0

BEGIN
NETWORK
TITLE =



NETWORK
TITLE =

      OPN   "DB LAUER";

NETWORK
TITLE =

      L     "MW 150";
      L     2#1011111110000000;
      AW    ;
      T     "MW 150";
      L     "MW 152";
      L     2#1111111111000000;
      AW    ;
      T     "MW 152";
NETWORK
TITLE =

      L     "MW 150";
      L     W#16#0;
      <>I   ;
      JC    M001;
      L     W#16#0;
      T     DBB   32;
M001: NOP   0;
NETWORK
TITLE =

      OPN   "DB LAUER";
      L     DBW    8;
      L     "MW 160";
      XOW   ;
      L     DBW    8;
      AW    ;
      T     "MW 162";
      TAK   ;
      L     "MW 160";
      AW    ;
      T     MW   164;
      L     DBW    8;
      T     "MW 160";
NETWORK
TITLE =

      OPN   "DB LAUER";
      L     DBW   10;
      L     "MW 170";
      XOW   ;
      L     DBW   10;
      AW    ;
      T     "MW 172";
      TAK   ;
      L     "MW 170";
      AW    ;
      T     MW   174;
      L     DBW   10;
      T     "MW 170";
NETWORK
TITLE =

      L     "MW 150";
      L     "MW 162";
      XOW   ;
      T     "MW 150";
NETWORK
TITLE =

      L     2#1011111110111111;
      L     "MW 150";
      AW    ;
      T     "MW 150";
NETWORK
TITLE =

      L     "MW 152";
      L     "MW 172";
      XOW   ;
      T     "MW 152";
NETWORK
TITLE =

      L     "MW 152";
      L     2#1011011111111111;
      AW    ;
      T     "MW 152";
NETWORK
TITLE =temps de controle de lamps

      A     "M 153.6";
      L     S5T#5S;
      SF    "Timer 0";
      NOP   0;
      NOP   0;
      NOP   0;
      NOP   0;
NETWORK
TITLE =

      A     "Timer 0";
      R     "M 153.6";
NETWORK
TITLE =

      A     "Timer 0";
      JC    M002;
      L     2#0;
      T     DBW   42;
      T     DBW   50;
      T     DBW   54;
M002: NOP   0;
NETWORK
TITLE =

      L     "MW 150";
      L     2#1111111111000000;
      AW    ;
      T     DBW   40;
NETWORK
TITLE =

      L     "MW 152";
      L     2#1111111111000000;
      AW    ;
      T     DBW   48;
NETWORK
TITLE =

      AN    "Timer 0";
      JC    M004;
      L     2#1111111111001111;
      T     DBW   42;
      T     DBW   46;
      T     DBW   50;
      T     DBW   54;
      L     2#110000;
      T     DBW   48;
M004: NOP   0;
NETWORK
TITLE =

      A     "Timer 0";
      JC    M005;
      L     W#16#0;
      L     DBW   42;
      L     DBW   50;
      L     DBW   54;
M005: NOP   0;
NETWORK
TITLE =

      AN    "M 134.0";
      JC    M006;
      L     DBW   44;
      L     2#100000000000;
      OW    ;
      T     DBW   44;
M006: NOP   0;
NETWORK
TITLE =

      AN    "M 134.2";
      JC    M007;
      L     DBW   44;
      L     2#1111011111111111;
      AW    ;
      T     DBW   44;
M007: NOP   0;
NETWORK
TITLE =
// BLD 131;
      O     "M 141.1";
      O     "M 141.2";
      O     "M 141.3";
      O     "M 141.4";
      O     "M 141.5";
      JC    M008;
      L     W#16#0;
      T     DBW   46;
      BEU   ;
M008: L     W#16#400;
      T     DBW   46;
NETWORK
TITLE =



END_FUNCTION

FUNCTION "LAUER SERVICE" : VOID
TITLE =Lauer Service
NAME : SERVICE
VERSION : 0.0

BEGIN
NETWORK
TITLE =

      OPN   "DB LAUER";

NETWORK
TITLE =

      AN    "M 150.5";
      JC    M001;
      L     DBW   72;
      L     2#100000000;
      T     DBW   72;
M001: NOP   0;
NETWORK
TITLE =

      AN    "M 150.5";
      JC    M002;
      L     2#11;
      T     DBW   76;
M002: NOP   0;
NETWORK
TITLE =

      AN    "M 150.5";
      JC    M003;
      A(    ;
      O     "M 161.0";
      O     "M 161.1";
      )     ;
      JC    M004;
      JU    M003;
M004: L     2#1000;
      T     DBB   74;
      JU    M005;
M003: L     DBB   74;
      L     2#11110111;
      AW    ;
      T     DBB   74;
M005: NOP   0;
NETWORK
TITLE =

      L     DBW   44;
      T     DBW   44;
NETWORK
TITLE =

      L     W#16#0;
      T     "MW 190";
NETWORK
TITLE =

      AN    "M 150.5";
      BEC   ;
NETWORK
TITLE =Service Mode - Elevator

      A(    ;
      L     DBB   32;
      L     1;
      <>I   ;
      )     ;
      JC    M006;
      =     "M 190.0";
      BEC   ;
M006: NOP   0;
NETWORK
TITLE =Service Mode - Flipper

      A(    ;
      L     DBB   32;
      L     2;
      <>I   ;
      )     ;
      JC    M007;
      =     "M 190.1";
      BEC   ;
M007: NOP   0;
NETWORK
TITLE =Service Mode - TurnTable

      A(    ;
      L     DBB   32;
      L     3;
      <>I   ;
      )     ;
      JC    M008;
      =     "M 190.2";
      BEC   ;
M008: NOP   0;
NETWORK
TITLE =

      A(    ;
      L     DBB   32;
      L     4;
      <>I   ;
      )     ;
      JC    M009;
      =     "M 190.3";
      BEC   ;
M009: NOP   0;
NETWORK
TITLE =

      A(    ;
      L     DBB   32;
      L     5;
      <>I   ;
      )     ;
      JC    M010;
      =     "M 190.4";
      BEC   ;
M010: NOP   0;
NETWORK
TITLE =

      A(    ;
      L     DBB   32;
      L     6;
      <>I   ;
      )     ;
      JC    M011;
      =     "M 190.5";
      BEC   ;
M011: NOP   0;
NETWORK
TITLE =

      A(    ;
      L     DBB   32;
      L     7;
      <>I   ;
      )     ;
      JC    M012;
      =     "M 190.6";
      BEC   ;
M012: NOP   0;
NETWORK
TITLE =

      A(    ;
      L     DBB   32;
      L     8;
      <>I   ;
      )     ;
      JC    M013;
      =     "M 190.7";
      BEC   ;
M013: NOP   0;
END_FUNCTION

FUNCTION "LAUER KEYS 2" : VOID
TITLE =Lauer Keys 2
NAME : ZEITEN1
VERSION : 0.0

BEGIN
NETWORK
TITLE =

      OPN   "DB LAUER";

NETWORK
TITLE =

      A     "M 171.0";
      BEC   ;
NETWORK
TITLE =

      AN    "M 151.7";
      JC    M001;
      L     2#100000000;
      T     DBW   72;
M001: NOP   0;
NETWORK
TITLE =

      AN    "M 151.7";
      JC    M002;
      L     2#1001;
      T     DBW   76;
M002: NOP   0;
NETWORK
TITLE =

      A     "M 171.0";
      BEC   ;
NETWORK
TITLE =

      A(    ;
      L     DBB   32;
      L     1;
      ==I   ;
      )     ;
      A     "M 151.7";
      JC    M003;
      JU    M003;

M003: CALL "LAUER TIME" (
           QUEL                     := DBW  240,
           _TIME                    := MW   130);


END_FUNCTION

FUNCTION "LAUER KEYS 3" : VOID
TITLE =Lauer Keys 3
//
NAME : _TIMER
VERSION : 0.0

BEGIN
NETWORK
TITLE =

      OPN   "DB LAUER";

NETWORK
TITLE =

      AN    "M 171.0";
      BEC   ;
NETWORK
TITLE =

      AN    "M 151.7";
      JC    M001;
      L     2#100000000;
      T     DBW   72;
M001: NOP   0;
NETWORK
TITLE =

      AN    "M 151.7";
      JC    M002;
      L     2#1011;
      T     DBW   76;
M002: NOP   0;
NETWORK
TITLE =

      A(    ;
      L     DBB   32;
      L     1;
      ==I   ;
      )     ;
      A     "M 151.7";
      JC    M003;
      JU    M004;
M003: JCN   X000;

      CALL "LAUER TIME" (
           QUEL                     := DBW  242,
           _TIME                    := MW   122);

X000: NOP   0;
M004: NOP   0;
NETWORK
TITLE =

      A(    ;
      L     DBB   32;
      L     2;
      ==I   ;
      )     ;
      A     "M 151.7";
      JC    M005;
      JU    M006;
M005: JCN   X001;

      CALL "LAUER TIME" (
           QUEL                     := DBW  252,
           _TIME                    := MW   124);

X001: NOP   0;
M006: NOP   0;
END_FUNCTION

FUNCTION "LAUER MESSAGE1" : VOID
TITLE =Faults
NAME : FEHLER1
VERSION : 0.0


VAR_TEMP
  MESSAGE_CUE : BOOL ;
END_VAR
BEGIN
NETWORK
TITLE =MESSAGE CUE
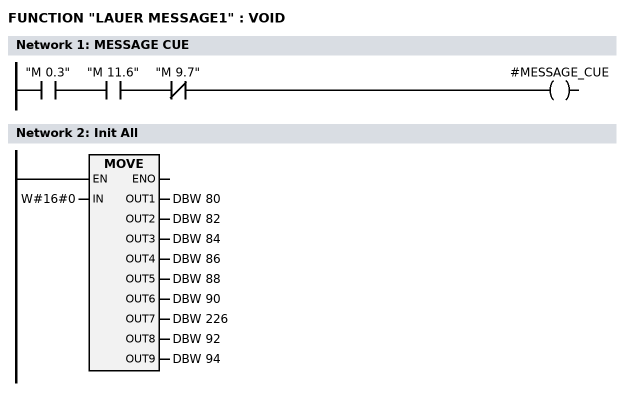

      A     "M 0.3";
      A     "M 11.6";
      AN    "M 9.7";
      =     #MESSAGE_CUE;
NETWORK
TITLE =Init All

      L     W#16#0;
      T     DBW   80;
      T     DBW   82;
      T     DBW   84;
      T     DBW   86;
      T     DBW   88;
      T     DBW   90;
      T     DBW  226;
      T     DBW   92;
      T     DBW   94;
NETWORK
TITLE =

      A     "M 0.4";
      JC    M001;
      JU    M002;
M001: L     2#100000000000;
      T     DBW   82;
      BEC   ;
M002: NOP   0;
NETWORK
TITLE =

      A     "M 22.7";
      JC    M003;
      JU    M004;
M003: L     2#1000;
      T     DBW   84;
      BEC   ;
M004: NOP   0;
NETWORK
TITLE =

      A     "M 1.0";
      JC    M005;
      JU    M006;
M005: L     2#10000;
      T     DBW   84;
      BEC   ;
M006: NOP   0;
NETWORK
TITLE =

      A     "M 1.1";
      JC    M007;
      JU    M008;
M007: L     2#100000;
      T     DBW   84;
      BEC   ;
M008: NOP   0;
NETWORK
TITLE =

      A     "M 1.2";
      JC    M009;
      JU    M010;
M009: L     2#1000000;
      T     DBW   84;
      BEC   ;
M010: NOP   0;
NETWORK
TITLE =

// Ancien alarme arrêt urgence élévateur 3
// maintenant libre
//      A     "M 1.3"
//      AN    "M 1.3"
//      JC    M011
//      JU    M012
///: L     2#10000000
//      T     DBW   84
//      BEC
//M012: NOP   0
NETWORK
TITLE =

      A     "M 1.3";
      JC    M013;
      JU    M014;
M013: L     2#100000000;
      T     DBW   84;
      BEC   ;
M014: NOP   0;
NETWORK
TITLE =

//     A     "M 1.5"
//     JC    M015
//      JU    M016
//M015: L     2#1000000000
//      T     DBW   84
//      BEC
//M016: NOP   0
NETWORK
TITLE =

      A     "M 0.5";
      JC    M017;
      JU    M018;
M017: L     2#10000000000;
      T     DBW   82;
      BEC   ;
M018: NOP   0;
NETWORK
TITLE =

      A     "M 0.6";
      JC    M019;
      JU    M020;
M019: L     2#1000000000000;
      T     DBW   82;
//;
      L     "MW 180";
      T     DBW  228;
      T     DBW  230;
      BEC   ;
M020: NOP   0;
NETWORK
TITLE =

      A     "M 0.7";
      JC    M021;
      JU    M022;
M021: L     2#10000000000000;
      T     DBW   82;
      BEC   ;
M022: NOP   0;
NETWORK
TITLE =

      O     "M 1.5";
      JC    M023;
      JU    M024;
M023: L     2#1;
      T     DBW   86;
      BEC   ;
M024: NOP   0;
NETWORK
TITLE =

      O     "M 30.1";
      JC    M025;
      JU    M026;
M025: L     2#10;
      T     DBW   86;
      BEC   ;
M026: NOP   0;
NETWORK
TITLE =

      O     "M 30.2";
      JC    M027;
      JU    M028;
M027: L     2#100;
      T     DBW   86;
      BEC   ;
M028: NOP   0;
NETWORK
TITLE =

      A     "M 1.6";
      JC    M029;
      JU    M030;
M029: L     2#100000000000000;
      T     DBW   84;
      BEC   ;
M030: NOP   0;
NETWORK
TITLE =

      A     "M 1.7";
      JC    M031;
      JU    M032;
M031: L     2#1000000000000000;
      T     DBW   84;
      BEC   ;
M032: NOP   0;
NETWORK
TITLE =

      A     "M 30.7";
      JC    M033;
      JU    M034;
M033: L     2#1000;
      T     DBW   86;
      BEC   ;
M034: NOP   0;
NETWORK
TITLE =

      A     "M 38.7";
      JC    M035;
      JU    M036;
M035: L     2#10000;
      T     DBW   86;
      BEC   ;
M036: NOP   0;
NETWORK
TITLE =

      A     "M 54.7";
      JC    M037;
      JU    M038;
M037: L     2#100000;
      T     DBW   86;
      BEC   ;
M038: NOP   0;
NETWORK
TITLE =

      O     "M 66.7";
      O     "M 86.7";
      JC    M039;
      JC    M040;
M039: L     2#1000000;
      T     DBW   86;
      BEC   ;
M040: NOP   0;
NETWORK
TITLE =

      A     "M 30.0";
      JC    M041;
      JU    M042;
M041: L     2#100000000;
      T     DBW   86;
      BEC   ;
M042: NOP   0;
NETWORK
TITLE =

      A     "M 98.1";
      JC    M043;
      JU    M044;
M043: L     2#10000000;
      T     DBW   86;
      BEC   ;
M044: NOP   0;
NETWORK
TITLE =

      A     "M 14.7";
      JC    M045;
      JU    M046;
M045: L     2#1000000000;
      T     DBW   86;
      BEC   ;
M046: NOP   0;
NETWORK
TITLE =

      A     "M 42.7";
      JC    M047;
      JU    M048;
M047: L     2#10000000000;
      T     DBW   86;
      BEC   ;
M048: NOP   0;
NETWORK
TITLE =

      A     #MESSAGE_CUE;
      A     "B 5.1";
      JC    M049;
      JU    M050;
M049: L     2#100000000000;
      T     DBW   86;
      L     2#10;
      T     DBW  232;
      BEC   ;
M050: NOP   0;
NETWORK
TITLE =

      A     #MESSAGE_CUE;
      A     "B 5.2";
      JC    M051;
      JU    M052;
M051: L     2#1000000000000;
      T     DBW   86;
      L     2#10;
      T     DBW  232;
      BEC   ;
M052: NOP   0;
NETWORK
TITLE =

      A     #MESSAGE_CUE;
      A     "B 5.4";
      JC    M053;
      JU    M054;
M053: L     2#10000000000000;
      T     DBW   86;
      L     2#10;
      T     DBW  232;
      BEC   ;
M054: NOP   0;
NETWORK
TITLE =

      A     #MESSAGE_CUE;
      A     "B 5.5";
      JC    M055;
      JU    M056;
M055: L     2#100000000000000;
      T     DBW   86;
      L     2#10;
      T     DBW  232;
      BEC   ;
M056: NOP   0;
NETWORK
TITLE =

      A     #MESSAGE_CUE;
      A     "B 6.0";
      JC    M057;
      JU    M058;
M057: L     2#1000000000000000;
      T     DBW   86;
      L     2#10;
      T     DBW  232;
      BEC   ;
M058: NOP   0;
NETWORK
TITLE =

      A     #MESSAGE_CUE;
      A     "B 6.7";
      O     "M 33.7";
      JC    M059;
      JU    M060;
M059: L     2#1;
      T     DBW   88;
      L     2#10;
      T     DBW  232;
      BEC   ;
M060: NOP   0;
NETWORK
TITLE =

      A     #MESSAGE_CUE;
      A     "B 7.0";
      JC    M061;
      JU    M062;
M061: L     2#10;
      T     DBW   88;
      L     2#10;
      T     DBW  232;
      BEC   ;
M062: NOP   0;
NETWORK
TITLE =

      A     #MESSAGE_CUE;
      A     "B 7.1";
      JC    M063;
      JU    M064;
M063: L     2#100;
      T     DBW   88;
      L     2#10;
      T     DBW  232;
      BEC   ;
M064: NOP   0;
NETWORK
TITLE =

      A     #MESSAGE_CUE;
      A     "B 7.2";
      JC    M065;
      JU    M066;
M065: L     2#1000;
      T     DBW   88;
      L     2#10;
      T     DBW  232;
      BEC   ;
M066: NOP   0;
NETWORK
TITLE =

      A     #MESSAGE_CUE;
      A     "B 7.3";
      JC    M067;
      JU    M068;
M067: L     2#10000;
      T     DBW   88;
      L     2#10;
      T     DBW  232;
      BEC   ;
M068: NOP   0;
NETWORK
TITLE =

      A     #MESSAGE_CUE;
      A     "B 7.4";
      JC    M069;
      JU    M070;
M069: L     2#100000;
      T     DBW   88;
      L     2#10;
      T     DBW  232;
      BEC   ;
M070: NOP   0;
NETWORK
TITLE =

      A     "M 98.2";
      JC    M071;
      JU    M072;
M071: L     2#1000000;
      T     DBW   88;
      BEC   ;
M072: NOP   0;
NETWORK
TITLE =

      A     #MESSAGE_CUE;
      A     "B 8.2";
      JC    M073;
      JU    M074;
M073: L     2#10000000;
      T     DBW   88;
      L     2#10;
      T     DBW  232;
      BEC   ;
M074: NOP   0;
NETWORK
TITLE =

      A     #MESSAGE_CUE;
      A     "B 9.6";
      JC    M075;
      JU    M076;
M075: L     2#100000000;
      T     DBW   88;
      L     2#10;
      T     DBW  232;
      BEC   ;
M076: NOP   0;
NETWORK
TITLE =

      A     #MESSAGE_CUE;
      A     "B 9.7";
      JC    M077;
      JU    M078;
M077: L     2#1000000000;
      T     DBW   88;
      L     2#10;
      T     DBW  232;
      BEC   ;
M078: NOP   0;
NETWORK
TITLE =

      A     #MESSAGE_CUE;
      A     "B 10.4";
      JC    M079;
      JU    M080;
M079: L     2#10000000000;
      T     DBW   88;
      L     2#10;
      T     DBW  232;
      BEC   ;
M080: NOP   0;
NETWORK
TITLE =

      A     #MESSAGE_CUE;
      A     "B 10.5";
      JC    M081;
      JU    M082;
M081: L     2#100000000000;
      T     DBW   88;
      L     2#10;
      T     DBW  232;
      BEC   ;
M082: NOP   0;
NETWORK
TITLE =

      A     #MESSAGE_CUE;
      A     "B 10.7";
      JC    M083;
      JU    M084;
M083: L     2#1000000000000;
      T     DBW   88;
      L     2#10;
      T     DBW  232;
      BEC   ;
M084: NOP   0;
NETWORK
TITLE =

      A     #MESSAGE_CUE;
      A     "B 11.0";
      JC    M085;
      JU    M086;
M085: L     2#10000000000000;
      T     DBW   88;
      L     2#10;
      T     DBW  232;
      BEC   ;
M086: NOP   0;
NETWORK
TITLE =

      A     #MESSAGE_CUE;
      A     "B 11.1";
      JC    M087;
      JU    M088;
M087: L     2#100000000000000;
      T     DBW   88;
      L     2#10;
      T     DBW  232;
      BEC   ;
M088: NOP   0;
NETWORK
TITLE =

//   A     #MESSAGE_CUE
//    AN    "B 11.1"
//     JC    M089
//     JU    M090
//M089: L     2#10
//      T     DBW   90
//      BEC
//M090: NOP   0
NETWORK
TITLE =

      A     #MESSAGE_CUE;
      AN    "B 5.4";
      JC    M091;
      JU    M092;
M091: L     2#100;
      T     DBW   90;
      BEC   ;
M092: NOP   0;
NETWORK
TITLE =

      A     #MESSAGE_CUE;
      AN    "B 9.7";
      JC    M093;
      JU    M094;
M093: L     2#1000;
      T     DBW   90;
      BEC   ;
M094: NOP   0;
NETWORK
TITLE =

      A     "M 11.7";
      JC    M095;
      JU    M096;
M095: L     2#1000000;
      T     DBW   90;
      BEC   ;
M096: NOP   0;
NETWORK
TITLE =

      A     "M 4.5";
      JC    M097;
      JU    M098;
M097: L     2#10000;
      T     DBW   90;
      L     1;
      T     DBW  226;
      BEC   ;
M098: NOP   0;
NETWORK
TITLE =

      A     "M 3.0";
      JC    M099;
      JU    M100;
M099: L     2#10000;
      T     DBW   90;
      L     2;
      T     DBW  226;
      BEC   ;
M100: NOP   0;
NETWORK
TITLE =

      A     "M 4.0";
      JC    M101;
      JU    M102;
M101: L     2#10000;
      T     DBW   90;
      L     3;
      T     DBW  226;
      BEC   ;
M102: NOP   0;
NETWORK
TITLE =

      A     "M 3.3";
      JC    M103;
      JU    M104;
M103: L     2#10000;
      T     DBW   90;
      L     4;
      T     DBW  226;
      BEC   ;
M104: NOP   0;
NETWORK
TITLE =

      A     "M 3.5";
      JC    M105;
      JU    M106;
M105: L     2#10000;
      T     DBW   90;
      L     5;
      T     DBW  226;
      BEC   ;
M106: NOP   0;
NETWORK
TITLE =

      A     "M 4.1";
      AN    "E 13.4";
      JC    M107;
      JU    M108;
M107: L     2#10000;
      T     DBW   90;
      L     6;
      T     DBW  226;
      BEC   ;
M108: NOP   0;
NETWORK
TITLE =

      A     "M 4.4";
      AN    "E 13.7";
      JC    M109;
      JU    M110;
M109: L     2#10000;
      T     DBW   90;
      L     7;
      T     DBW  226;
      BEC   ;
M110: NOP   0;
NETWORK
TITLE =

      A     "M 3.1";
      JC    M111;
      JU    M112;
M111: L     2#10000;
      T     DBW   90;
      L     8;
      T     DBW  226;
      BEC   ;
M112: NOP   0;
NETWORK
TITLE =

      A     "M 3.2";
      JC    M113;
      JU    M114;
M113: L     2#10000;
      T     DBW   90;
      L     9;
      T     DBW  226;
      BEC   ;
M114: NOP   0;
NETWORK
TITLE =

      A     "M 3.4";
      JC    M115;
      JU    M116;
M115: L     2#10000;
      T     DBW   90;
      L     10;
      T     DBW  226;
      BEC   ;
M116: NOP   0;
NETWORK
TITLE =

      A     "M 3.6";
      JC    M117;
      JU    M118;
M117: L     2#10000;
      T     DBW   90;
      L     11;
      T     DBW  226;
      BEC   ;
M118: NOP   0;
NETWORK
TITLE =

      A     "M 3.7";
      JC    M119;
      JU    M120;
M119: L     2#10000;
      T     DBW   90;
      L     12;
      T     DBW  226;
      BEC   ;
M120: NOP   0;
NETWORK
TITLE =

      A     "M 4.6";
      JC    M121;
      JU    M122;
M121: L     2#10000;
      T     DBW   90;
      L     13;
      T     DBW  226;
      BEC   ;
M122: NOP   0;
NETWORK
TITLE =

      A     "M 4.1";
      JC    M123;
      JU    M124;
M123: L     2#10000;
      T     DBW   90;
      L     14;
      T     DBW  226;
      BEC   ;
M124: NOP   0;
NETWORK
TITLE =

      A     "M 4.3";
      AN    "E 13.6";
      JC    M125;
      JU    M126;
M125: L     2#10000;
      T     DBW   90;
      L     15;
      T     DBW  226;
      BEC   ;
M126: NOP   0;
NETWORK
TITLE =

      A     "M 4.1";
      AN    "E 28.0";
      JC    M127;
      JU    M128;
M127: L     2#10000;
      T     DBW   90;
      L     16;
      T     DBW  226;
      BEC   ;
M128: NOP   0;
NETWORK
TITLE =

      A     "M 4.1";
      AN    "E 28.1";
      JC    M129;
      JU    M130;
M129: L     2#10000;
      T     DBW   90;
      L     17;
      T     DBW  226;
      BEC   ;
M130: NOP   0;
NETWORK
TITLE =

      A     "M 4.1";
      AN    "E 28.2";
      JC    M131;
      JU    M132;
M131: L     2#10000;
      T     DBW   90;
      L     18;
      T     DBW  226;
      BEC   ;
M132: NOP   0;
NETWORK
TITLE =

// Affichage d'alarme libéré de l'ancien 506
// maintenant libre
//      A     "M 0.3"
//      AN    "M 0.3"
//      JC    M133
//      JU    M134
//M133: L     2#10000
//      T     DBW   90
//      L     19
//      T     DBW  226
//      BEC
//M134: NOP   0
NETWORK
TITLE =

// Affichage d'alarme libéré de l'ancien 506
// maintenant libre
////      A     "M 0.3"
//      AN    "M 0.3"
//      JC    M135
//     JU    M136
//M135: L     2#10000
//      T     DBW   90
//      L     20
//      T     DBW  226
//      BEC
//M136: NOP   0
NETWORK
TITLE =

// Affichage d'alarme libéré de l'ancien 506
// maintenant libre
//     A     "M 0.3"
//     AN    "M 0.3"
//      JC    M137
//      JU    M138
//M137: L     2#10000
//      T     DBW   90
//      L     21
//      T     DBW  226
//      BEC
//M138: NOP   0
NETWORK
TITLE =

// Affichage d'alarme libéré de l'ancien 506
// maintenant libre
//      A     "M 0.3"
//      AN    "M 0.3"
//      JC    M139
//      JU    M140
//M139: L     2#10000
//      T     DBW   90
//      L     22
//      T     DBW  226
//      BEC
//M140: NOP   0
NETWORK
TITLE =

// Affichage d'alarme libéré de l'ancien 506
// maintenant libre
//     A     "M 0.3"
//     AN    "M 0.3"
//     JC    M141
//     JU    M142
//M141: L     2#10000
//      T     DBW   90
//      L     23
//      T     DBW  226
//      BEC
//M142: NOP   0
NETWORK
TITLE =

// Affichage d'alarme libéré de l'ancien 506
// maintenant libre
//      A     "M 0.3"
//      AN    "M 0.3"
//      JC    M143
//      JU    M144
//M143: L     2#10000
//      T     DBW   90
//      L     24
//      T     DBW  226
//      BEC
//M144: NOP   0
NETWORK
TITLE =

// Affichage d'alarme libéré de l'ancien 506
// maintenant libre
//      A     "M 0.3"
////      AN    "M 0.3"
//      JC    M145
//      JU    M146
//M145: L     2#10000
//      T     DBW   90
//      L     25
//      T     DBW  226
//      BEC
//M146: NOP   0
NETWORK
TITLE =

      A     "Timer 0";
      JC    M147;
      JC    M148;
M147: L     2#100000;
      T     DBW   94;
      BEC   ;
M148: NOP   0;
NETWORK
TITLE =

// Affichage d'alarme libéré de l'ancien 506
// maintenant libre
//      A     M      2.3
//      AN    M      2.3
//      JC    M149
//      JC    M150
//M149: L     2#1000
//     T     DBW   94
//     BEC
//M150: NOP   0
NETWORK
TITLE =

      O     "M 150.2";
      JC    M151;
      JC    M152;
M151: L     2#10000;
      T     DBW   94;
//;
      BEC   ;
M152: NOP   0;
NETWORK
TITLE =

      A     "M 10.0";
      JC    M153;
      JU    M154;
M153: L     2#10000000;
      T     DBW   90;
      BEC   ;
M154: NOP   0;
END_FUNCTION

FUNCTION "LAUER MESSAGE2" : VOID
TITLE =Lauer Message 2
NAME : STATUS
VERSION : 0.0

BEGIN
NETWORK
TITLE =

      OPN   "DB LAUER";

NETWORK
TITLE =

      A(    ;
      O     "M 150.4";
      O     "M 150.5";
      O     "M 150.7";
      ON    "S 2.1";
      O     "S 2.2";
      )     ;
      AN    "M 0.1";
      AN    "M 0.2";
      AN    "M 0.3";
      AN    "M 1.5";
      AN    "M 1.7";
//;
      JC    M001;
      JU    M002;
M001: L     2#100;
      T     DBW   82;
      BEC   ;
M002: NOP   0;
NETWORK
TITLE =

      A     "M 0.2";
      AN    "M 0.3";
      JC    M003;
      JU    M004;
M003: L     2#1000;
      T     DBW   82;
      BEC   ;
M004: NOP   0;
NETWORK
TITLE =

      A     "M 0.3";
      AN    "M 9.7";
      JC    M005;
      JU    M006;
M005: L     2#10000;
      T     DBW   82;
      BEC   ;
M006: NOP   0;
END_FUNCTION

FUNCTION "LAUER CALL" : VOID
TITLE =Lauer Call
// TEXT ORG
NAME : TEXTORG
VERSION : 0.0

BEGIN
NETWORK
TITLE =

      OPN   "DB LAUER";

NETWORK
TITLE =Reset & Preset
//When the communication/control byte is in a neutral state, and those two
//internal flags are off, the FC restores default preset values in the Lauer DB.
      A(    ;
      L     "MB 150";
      L     W#16#FFF7;
      AW    ;
      L     W#16#0;
      )     ;
      ==I   ;
      AN    "M 151.6";
      AN    "M 151.7";
      JC    M001;
      JU    M002;

M001: L     2#0;
      T     DBW   76;
//;
      L     2#111100000000;
      T     DBW   72;
//;
      L     2#11100000000001;
      T     DBW   74;
//;
      L     W#16#0;
      T     DBW   32;

M002: NOP   0;
NETWORK
TITLE =
//transfer keypad/page/request words
//avoid repeated copying every scan
//only copy
//once per trigger edge/state
      A     "M 0.3";
      AN    "M 200.0";
      JC    M003;
      A     "M 0.2";
      AN    "M 200.1";
      JC    M004;
      JU    M005;

M003: L     "MW 150";
      T     "MW 118";
//;
      L     "MW 152";
      T     "MW 120";
//;
      A     "M 0.3";
      S     "M 200.0";
      R     "M 200.1";
      JU    M005;

M004: L     "MW 118";
      T     "MW 150";
//;
      L     "MW 120";
      T     "MW 152";
//;
      A     "M 0.2";
      S     "M 200.1";
      R     "M 200.0";

M005: NOP   0;
NETWORK
TITLE =
//reopen "DB LAUER"
//
//load DBW48
//
//call LAUER KEYS 1
      OPN   "DB LAUER";
      L     DBW   48;
      CALL "LAUER KEYS 1" ;
NETWORK
TITLE =

      CALL "LAUER SERVICE" ;

NETWORK
TITLE =

      CALL "LAUER KEYS 2" ;

NETWORK
TITLE =

      CALL "LAUER KEYS 3" ;

NETWORK
TITLE =

      CALL "LAUER MESSAGE1" ;

NETWORK
TITLE =

//      CALL  "LAUER"

NETWORK
TITLE =

      CALL "LAUER MESSAGE2" ;

END_FUNCTION

FUNCTION "SETUP" : VOID
TITLE =Setup Values
//Do Not Change These Values !!!
NAME : SETUP
VERSION : 0.1

BEGIN
NETWORK
TITLE =Setup Values - Slat Conveyor 3

      L     8000;
      T     "COLLATORS DB".Conveyor_Length_C3;
NETWORK
TITLE =Setup Values - Conveyor 4

      L     800; //900
      T     "COLLATORS DB".Surface_Length_C4;
NETWORK
TITLE =Setup Value  - TurnTable - Need " Packet IN " to Start

      S     "M 47.4";

NETWORK
TITLE =Setup Values - Conveyor 10

      L     13000;
      T     "COLLATORS DB".Surface_Length_10;
NETWORK
TITLE =Counter Setup


      S     "M 167.7";
NETWORK
TITLE =Packet Counter Constants 11.0 & 5.5

      L     1.000000e+01;
      T     "DB UTILITY".LENGTH_CONST;
//;
      L     5.200000e-01;
      T     "DB UTILITY".WIDTH_CONST;
NETWORK
TITLE =HMI - Conveyor Time

      L     150;
      T     "HMI_DB".CONV_7_POS_mS;
//;
      L     30;
      T     "HMI_DB".CONV_8_POS_FWD_mS;
//;
      L     70;
      T     "HMI_DB".CONV_8_POS_REV_mS;
//;
      L     15;
      T     "HMI_DB".CONV_9_POS_mS;
NETWORK
TITLE =HMI Control - Reset

      R     "HMI_DB".ON_SW;
      R     "HMI_DB".SERVICE_SW_1_STATUS;
      R     "HMI_DB".SERVICE_SW_2_STATUS;
      R     "HMI_DB".SERVICE_SW_3_STATUS;
      R     "HMI_DB".SERVICE_SW_1_2_STATUS;
END_FUNCTION

FUNCTION "SENSOR DE-BOUNCER" : VOID
TITLE =Sensor Debouncer
//Counting Foul Sensor Switching of less than PreSet Time
VERSION : 0.2


VAR_INPUT
  Bit_0 : BOOL ;
  Bit_1 : BOOL ;
  Preset_mS : INT ;
  Debounce_mS : INT ;
  Plc_Scan_mS : INT ;
END_VAR
VAR_IN_OUT
  Rising_Pulse_1 : BOOL ;	//Db Struct
  Rising_Pulse_2 : BOOL ;	//Db Struct
  Rising_Pulse_3 : BOOL ;	//Db Struct
  Rising_Pulse_4 : BOOL ;	//Db Struct
  Rising_Pulse_5 : BOOL ;	//Db Struct
  Rising_Pulse_6 : BOOL ;	//Db Struct
  Rising_Pulse_7 : BOOL ;	//Db Struct
  Rising_Pulse_8 : BOOL ;	//Db Struct
  Memory_Bit_1 : BOOL ;	//Db Struct
  Memory_Bit_2 : BOOL ;	//Db Struct
  Memory_Bit_3 : BOOL ;	//Db Struct
  Memory_Bit_4 : BOOL ;	//Db Struct
  Memory_Bit_5 : BOOL ;	//Db Struct
  Memory_Bit_6 : BOOL ;	//Db Struct
  Spare_1 : BOOL ;	//Db Struct
  Spare_2 : BOOL ;	//Db Struct
  Word_Buffer_1 : INT ;	//Db Struct
  Word_Buffer_2 : INT ;	//Db Struct
  Word_Result : INT ;	//Db Struct
  Word_Count_Limit : INT ;	//Db Data
  Word_Count : INT ;	//Db/HMI Data
END_VAR
VAR_TEMP
  MEMORY_1 : BOOL ;
  MEMORY_2 : BOOL ;
  MEMORY_3 : BOOL ;
END_VAR
BEGIN
NETWORK
TITLE =Init on First Call

      A     #Memory_Bit_6;
      JNB   INI1;
      JU    INI2;

INI1: L     0;
      T     #Word_Buffer_1;
      T     #Word_Buffer_2;
      R     #Memory_Bit_1;
      R     #Memory_Bit_2;
      R     #Memory_Bit_3;
      R     #Memory_Bit_4;
      R     #Memory_Bit_5;
      S     #Memory_Bit_6;

INI2: NOP   0;

NETWORK
TITLE =Input Bits - Start Event
//- #Bit_0 : Conveyor X InFeed Sensor
//- #Bit_1 : Conveyor X Exit Sensor
      A     #Bit_0;
      FP    #Rising_Pulse_1;
      JNB   K001;
      L     0;
      T     #Word_Buffer_1;
      R     #Memory_Bit_4;
      S     #Memory_Bit_1;

K001: NOP   0;

      A     #Bit_1;
      FP    #Rising_Pulse_2;
      JNB   K002;
      L     0;
      T     #Word_Buffer_2;
      S     #Memory_Bit_2;

K002: NOP   0;

NETWORK
TITLE =TimeBase
//TimeBase -> ScanTime
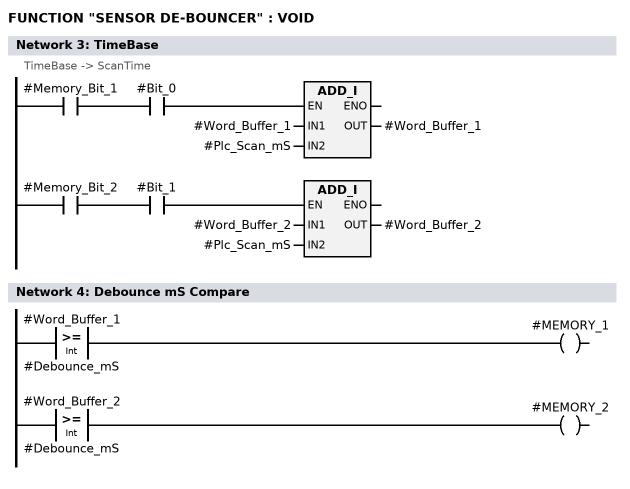
      A     #Memory_Bit_1;
      A     #Bit_0;
      JNB   K003;
      L     #Word_Buffer_1;
      L     #Plc_Scan_mS;
      +I    ;
      T     #Word_Buffer_1;

K003: NOP   0;

      A     #Memory_Bit_2;
      A     #Bit_1;
      JNB   K004;
      L     #Word_Buffer_2;
      L     #Plc_Scan_mS;
      +I    ;
      T     #Word_Buffer_2;

K004: NOP   0;

NETWORK
TITLE =Debounce mS Compare

      A(    ;
      L     #Word_Buffer_1;
      L     #Debounce_mS;
      >=I   ;
      )     ;
      =     #MEMORY_1;
//;
      A(    ;
      L     #Word_Buffer_2;
      L     #Debounce_mS;
      >=I   ;
      )     ;
      =     #MEMORY_2;

NETWORK
TITLE =Add to Packet Number with Bit_0
//Validated ON event on Bit_0 adds +1 one time
      A     #Memory_Bit_1;
      A     #MEMORY_1;
      A     #Bit_0;
      FP    #Rising_Pulse_4;
      JNB   K005;
      L     #Word_Count;
      L     1;
      +I    ;
      T     #Word_Count;
      R     #Memory_Bit_1;

K005: NOP   0;

NETWORK
TITLE =Subtract from Packet Number with Bit_1
//Validated ON event on Bit_1 subtracts -1 on falling edge
      AN    #Bit_1;
      FP    #Rising_Pulse_5;
      JNB   K006;

      A     #Memory_Bit_2;
      A     #MEMORY_2;
      JNB   K006;
//;
      L     #Word_Count;
      L     1;
      -I    ;
      T     #Word_Count;
      R     #Memory_Bit_2;

K006: NOP   0;

NETWORK
TITLE =Clamp Packet Number
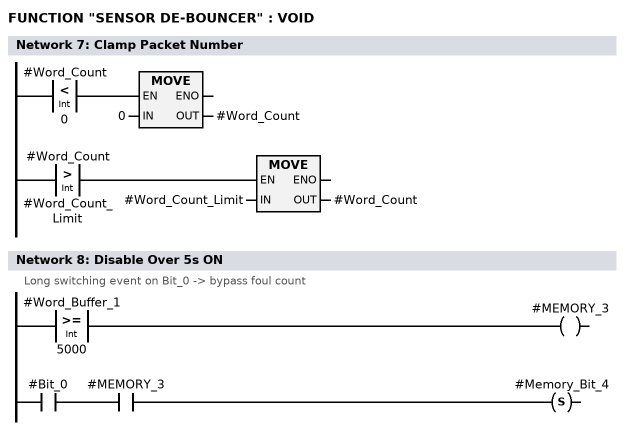

      L     #Word_Count;
      L     0;
      <I    ;
      JNB   K007;
      L     0;
      T     #Word_Count;

K007: NOP   0;

      L     #Word_Count;
      L     #Word_Count_Limit;
      >I    ;
      JNB   K008;
      L     #Word_Count_Limit;
      T     #Word_Count;

K008: NOP   0;

NETWORK
TITLE =Disable Over 5s ON
//Long switching event on Bit_0 -> bypass foul count
      L     #Word_Buffer_1;
      L     5000;
      >=I   ;
      =     #MEMORY_3;
//;
      A     #Bit_0;
      A     #MEMORY_3;
      S     #Memory_Bit_4;

NETWORK
TITLE =Result
//Word_Result +1 if Bit_0 turns OFF before Preset_mS and was not bypassed
      AN    #Bit_0;
      FP    #Rising_Pulse_6;
      JNB   K009;

      A     #Memory_Bit_1;
      AN    #Memory_Bit_4;
      JNB   K010;
//;
      L     #Word_Buffer_1;
      L     #Preset_mS;
      <I    ;
      JNB   K010;
//;
      L     #Word_Result;
      L     1;
      +I    ;
      T     #Word_Result;

K010: R     #Memory_Bit_1;
      R     #Memory_Bit_4;
      L     0;
      T     #Word_Buffer_1;

K009: NOP   0;

NETWORK
TITLE =Reset Exit Event on Falling Edge

      AN    #Bit_1;
      FP    #Rising_Pulse_7;
      JNB   K011;
      R     #Memory_Bit_2;
      L     0;
      T     #Word_Buffer_2;

K011: NOP   0;

END_FUNCTION

FUNCTION "SENSOR CHECK CALLS" : VOID
TITLE =
VERSION : 0.1

BEGIN
NETWORK
TITLE =
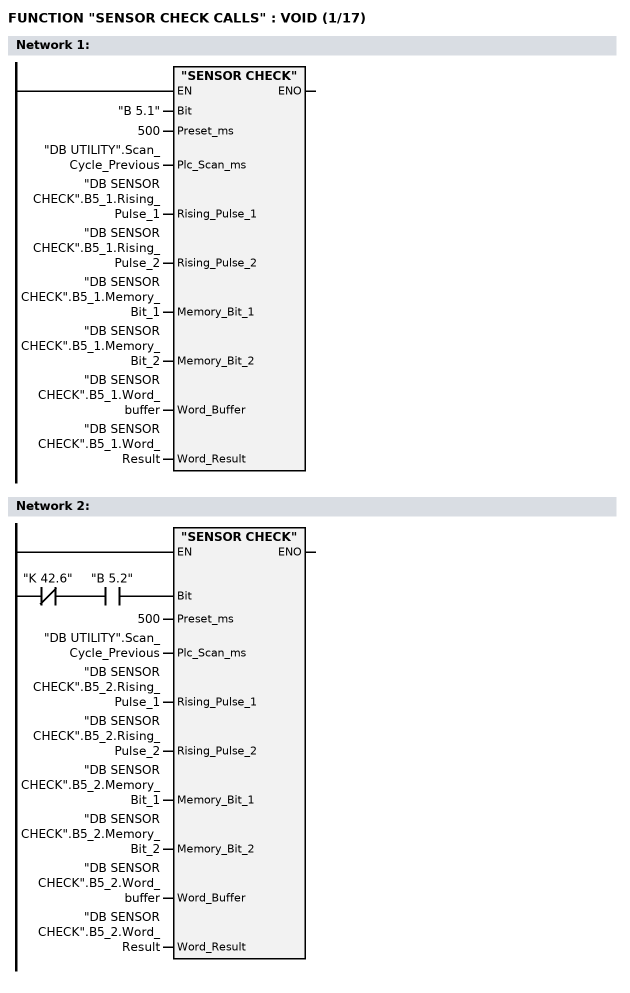

      CALL "SENSOR CHECK" (
           Bit                      := "B 5.1",
           Preset_ms                := 500,
           Plc_Scan_ms              := "DB UTILITY".Scan_Cycle_Previous,
           Rising_Pulse_1           := "DB SENSOR CHECK".B5_1.Rising_Pulse_1,
           Rising_Pulse_2           := "DB SENSOR CHECK".B5_1.Rising_Pulse_2,
           Memory_Bit_1             := "DB SENSOR CHECK".B5_1.Memory_Bit_1,
           Memory_Bit_2             := "DB SENSOR CHECK".B5_1.Memory_Bit_2,
           Word_Buffer              := "DB SENSOR CHECK".B5_1.Word_buffer,
           Word_Result              := "DB SENSOR CHECK".B5_1.Word_Result);

NETWORK
TITLE =

      AN    "K 42.6";
      A     "B 5.2";
      =     L      0.0;
//;
      CALL "SENSOR CHECK" (
           Bit                      := L      0.0,
           Preset_ms                := 500,
           Plc_Scan_ms              := "DB UTILITY".Scan_Cycle_Previous,
           Rising_Pulse_1           := "DB SENSOR CHECK".B5_2.Rising_Pulse_1,
           Rising_Pulse_2           := "DB SENSOR CHECK".B5_2.Rising_Pulse_2,
           Memory_Bit_1             := "DB SENSOR CHECK".B5_2.Memory_Bit_1,
           Memory_Bit_2             := "DB SENSOR CHECK".B5_2.Memory_Bit_2,
           Word_Buffer              := "DB SENSOR CHECK".B5_2.Word_buffer,
           Word_Result              := "DB SENSOR CHECK".B5_2.Word_Result);

NETWORK
TITLE =
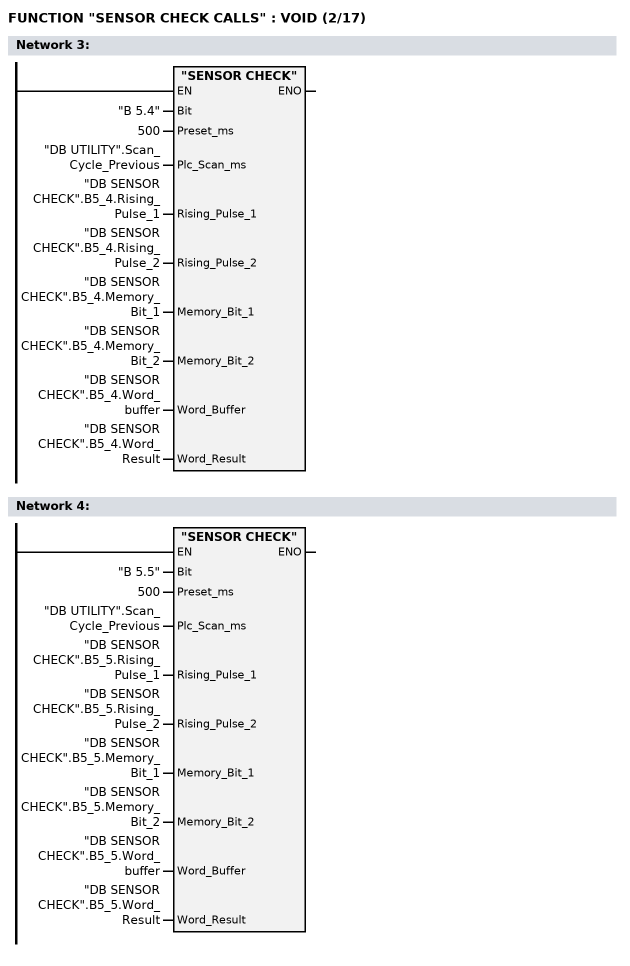

      CALL "SENSOR CHECK" (
           Bit                      := "B 5.4",
           Preset_ms                := 500,
           Plc_Scan_ms              := "DB UTILITY".Scan_Cycle_Previous,
           Rising_Pulse_1           := "DB SENSOR CHECK".B5_4.Rising_Pulse_1,
           Rising_Pulse_2           := "DB SENSOR CHECK".B5_4.Rising_Pulse_2,
           Memory_Bit_1             := "DB SENSOR CHECK".B5_4.Memory_Bit_1,
           Memory_Bit_2             := "DB SENSOR CHECK".B5_4.Memory_Bit_2,
           Word_Buffer              := "DB SENSOR CHECK".B5_4.Word_buffer,
           Word_Result              := "DB SENSOR CHECK".B5_4.Word_Result);

NETWORK
TITLE =

      CALL "SENSOR CHECK" (
           Bit                      := "B 5.5",
           Preset_ms                := 500,
           Plc_Scan_ms              := "DB UTILITY".Scan_Cycle_Previous,
           Rising_Pulse_1           := "DB SENSOR CHECK".B5_5.Rising_Pulse_1,
           Rising_Pulse_2           := "DB SENSOR CHECK".B5_5.Rising_Pulse_2,
           Memory_Bit_1             := "DB SENSOR CHECK".B5_5.Memory_Bit_1,
           Memory_Bit_2             := "DB SENSOR CHECK".B5_5.Memory_Bit_2,
           Word_Buffer              := "DB SENSOR CHECK".B5_5.Word_buffer,
           Word_Result              := "DB SENSOR CHECK".B5_5.Word_Result);

NETWORK
TITLE =
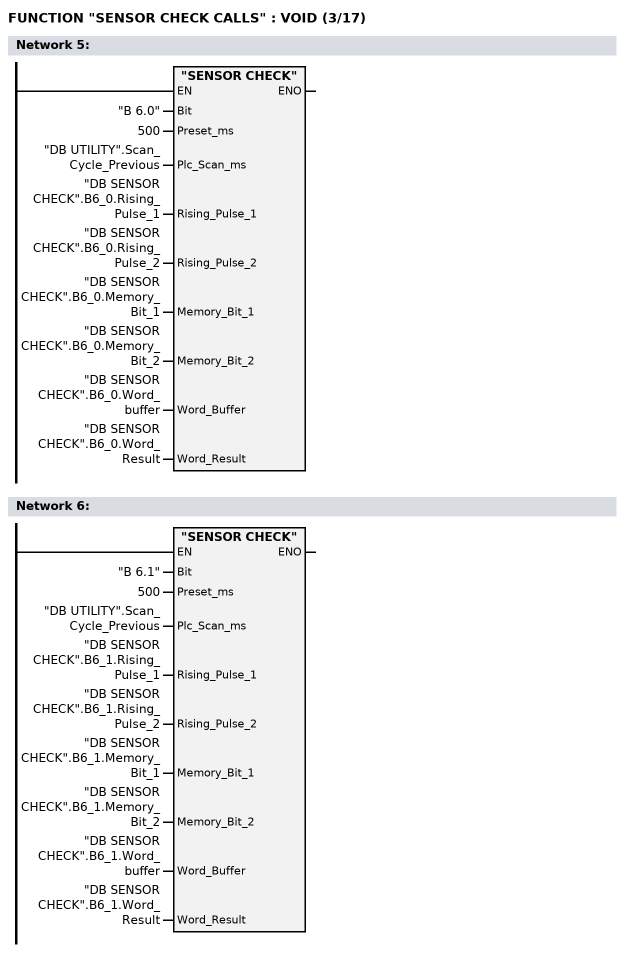

      CALL "SENSOR CHECK" (
           Bit                      := "B 6.0",
           Preset_ms                := 500,
           Plc_Scan_ms              := "DB UTILITY".Scan_Cycle_Previous,
           Rising_Pulse_1           := "DB SENSOR CHECK".B6_0.Rising_Pulse_1,
           Rising_Pulse_2           := "DB SENSOR CHECK".B6_0.Rising_Pulse_2,
           Memory_Bit_1             := "DB SENSOR CHECK".B6_0.Memory_Bit_1,
           Memory_Bit_2             := "DB SENSOR CHECK".B6_0.Memory_Bit_2,
           Word_Buffer              := "DB SENSOR CHECK".B6_0.Word_buffer,
           Word_Result              := "DB SENSOR CHECK".B6_0.Word_Result);

NETWORK
TITLE =

      CALL "SENSOR CHECK" (
           Bit                      := "B 6.1",
           Preset_ms                := 500,
           Plc_Scan_ms              := "DB UTILITY".Scan_Cycle_Previous,
           Rising_Pulse_1           := "DB SENSOR CHECK".B6_1.Rising_Pulse_1,
           Rising_Pulse_2           := "DB SENSOR CHECK".B6_1.Rising_Pulse_2,
           Memory_Bit_1             := "DB SENSOR CHECK".B6_1.Memory_Bit_1,
           Memory_Bit_2             := "DB SENSOR CHECK".B6_1.Memory_Bit_2,
           Word_Buffer              := "DB SENSOR CHECK".B6_1.Word_buffer,
           Word_Result              := "DB SENSOR CHECK".B6_1.Word_Result);

NETWORK
TITLE =
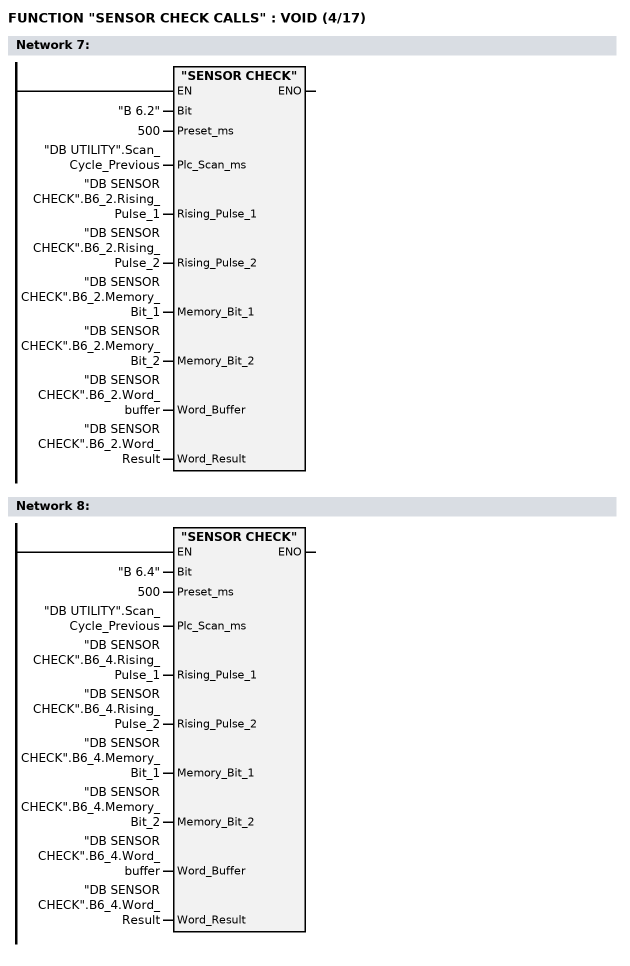

      CALL "SENSOR CHECK" (
           Bit                      := "B 6.2",
           Preset_ms                := 500,
           Plc_Scan_ms              := "DB UTILITY".Scan_Cycle_Previous,
           Rising_Pulse_1           := "DB SENSOR CHECK".B6_2.Rising_Pulse_1,
           Rising_Pulse_2           := "DB SENSOR CHECK".B6_2.Rising_Pulse_2,
           Memory_Bit_1             := "DB SENSOR CHECK".B6_2.Memory_Bit_1,
           Memory_Bit_2             := "DB SENSOR CHECK".B6_2.Memory_Bit_2,
           Word_Buffer              := "DB SENSOR CHECK".B6_2.Word_buffer,
           Word_Result              := "DB SENSOR CHECK".B6_2.Word_Result);

NETWORK
TITLE =

      CALL "SENSOR CHECK" (
           Bit                      := "B 6.4",
           Preset_ms                := 500,
           Plc_Scan_ms              := "DB UTILITY".Scan_Cycle_Previous,
           Rising_Pulse_1           := "DB SENSOR CHECK".B6_4.Rising_Pulse_1,
           Rising_Pulse_2           := "DB SENSOR CHECK".B6_4.Rising_Pulse_2,
           Memory_Bit_1             := "DB SENSOR CHECK".B6_4.Memory_Bit_1,
           Memory_Bit_2             := "DB SENSOR CHECK".B6_4.Memory_Bit_2,
           Word_Buffer              := "DB SENSOR CHECK".B6_4.Word_buffer,
           Word_Result              := "DB SENSOR CHECK".B6_4.Word_Result);

NETWORK
TITLE =
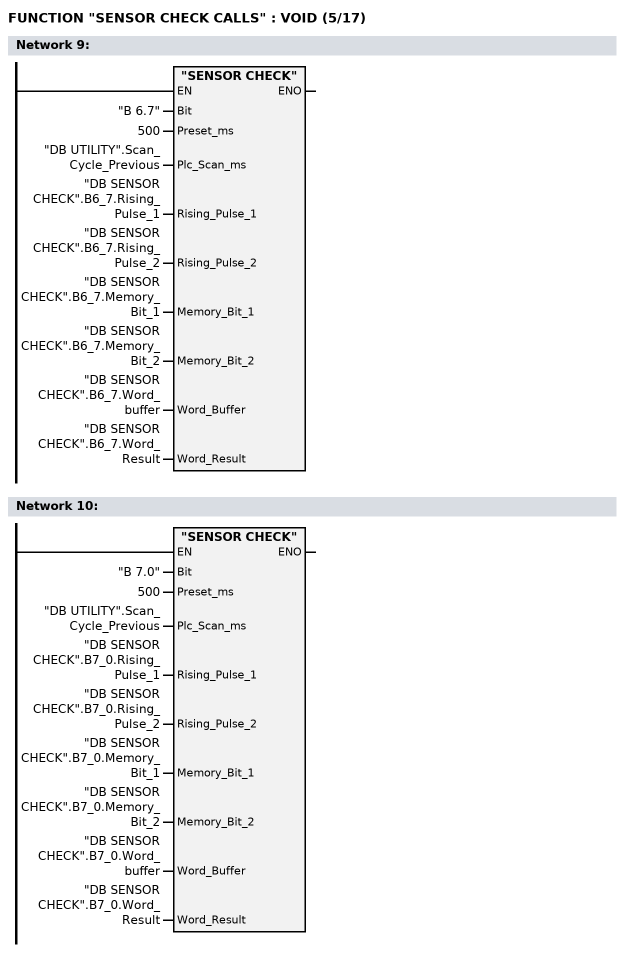

      CALL "SENSOR CHECK" (
           Bit                      := "B 6.7",
           Preset_ms                := 500,
           Plc_Scan_ms              := "DB UTILITY".Scan_Cycle_Previous,
           Rising_Pulse_1           := "DB SENSOR CHECK".B6_7.Rising_Pulse_1,
           Rising_Pulse_2           := "DB SENSOR CHECK".B6_7.Rising_Pulse_2,
           Memory_Bit_1             := "DB SENSOR CHECK".B6_7.Memory_Bit_1,
           Memory_Bit_2             := "DB SENSOR CHECK".B6_7.Memory_Bit_2,
           Word_Buffer              := "DB SENSOR CHECK".B6_7.Word_buffer,
           Word_Result              := "DB SENSOR CHECK".B6_7.Word_Result);

NETWORK
TITLE =

      CALL "SENSOR CHECK" (
           Bit                      := "B 7.0",
           Preset_ms                := 500,
           Plc_Scan_ms              := "DB UTILITY".Scan_Cycle_Previous,
           Rising_Pulse_1           := "DB SENSOR CHECK".B7_0.Rising_Pulse_1,
           Rising_Pulse_2           := "DB SENSOR CHECK".B7_0.Rising_Pulse_2,
           Memory_Bit_1             := "DB SENSOR CHECK".B7_0.Memory_Bit_1,
           Memory_Bit_2             := "DB SENSOR CHECK".B7_0.Memory_Bit_2,
           Word_Buffer              := "DB SENSOR CHECK".B7_0.Word_buffer,
           Word_Result              := "DB SENSOR CHECK".B7_0.Word_Result);

NETWORK
TITLE =
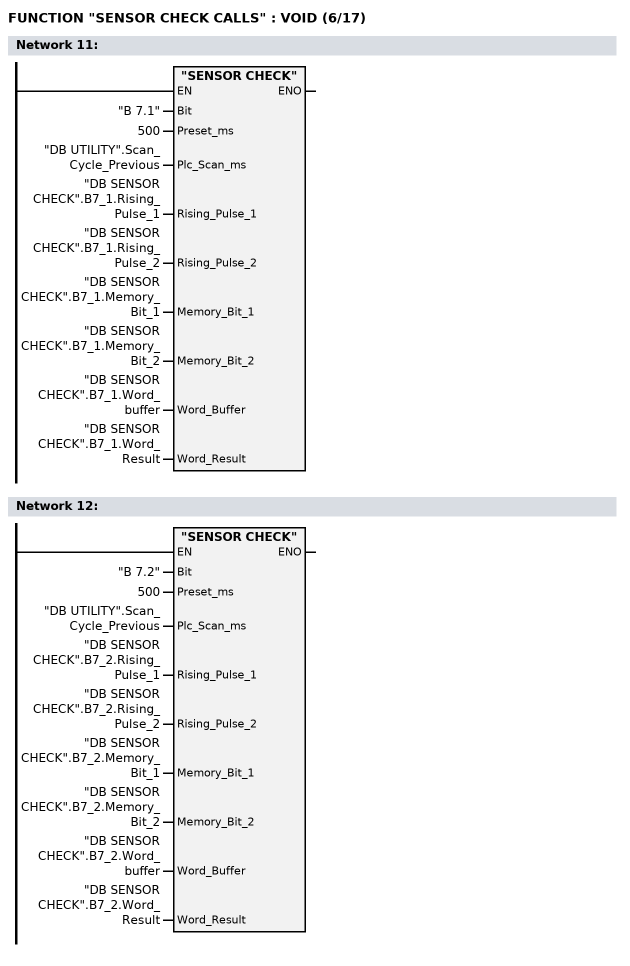

      CALL "SENSOR CHECK" (
           Bit                      := "B 7.1",
           Preset_ms                := 500,
           Plc_Scan_ms              := "DB UTILITY".Scan_Cycle_Previous,
           Rising_Pulse_1           := "DB SENSOR CHECK".B7_1.Rising_Pulse_1,
           Rising_Pulse_2           := "DB SENSOR CHECK".B7_1.Rising_Pulse_2,
           Memory_Bit_1             := "DB SENSOR CHECK".B7_1.Memory_Bit_1,
           Memory_Bit_2             := "DB SENSOR CHECK".B7_1.Memory_Bit_2,
           Word_Buffer              := "DB SENSOR CHECK".B7_1.Word_buffer,
           Word_Result              := "DB SENSOR CHECK".B7_1.Word_Result);

NETWORK
TITLE =

      CALL "SENSOR CHECK" (
           Bit                      := "B 7.2",
           Preset_ms                := 500,
           Plc_Scan_ms              := "DB UTILITY".Scan_Cycle_Previous,
           Rising_Pulse_1           := "DB SENSOR CHECK".B7_2.Rising_Pulse_1,
           Rising_Pulse_2           := "DB SENSOR CHECK".B7_2.Rising_Pulse_2,
           Memory_Bit_1             := "DB SENSOR CHECK".B7_2.Memory_Bit_1,
           Memory_Bit_2             := "DB SENSOR CHECK".B7_2.Memory_Bit_2,
           Word_Buffer              := "DB SENSOR CHECK".B7_2.Word_buffer,
           Word_Result              := "DB SENSOR CHECK".B7_2.Word_Result);

NETWORK
TITLE =
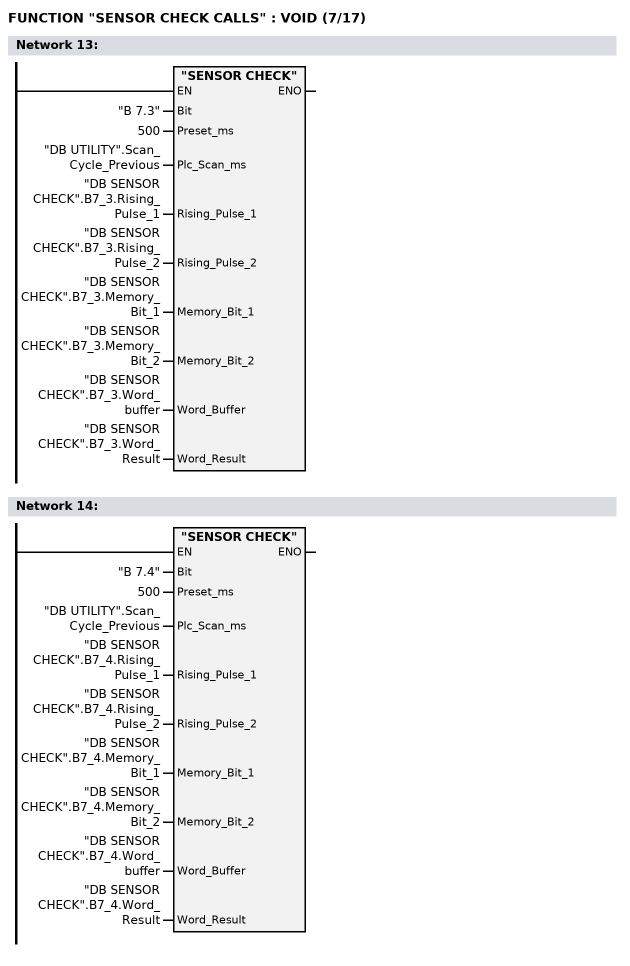

      CALL "SENSOR CHECK" (
           Bit                      := "B 7.3",
           Preset_ms                := 500,
           Plc_Scan_ms              := "DB UTILITY".Scan_Cycle_Previous,
           Rising_Pulse_1           := "DB SENSOR CHECK".B7_3.Rising_Pulse_1,
           Rising_Pulse_2           := "DB SENSOR CHECK".B7_3.Rising_Pulse_2,
           Memory_Bit_1             := "DB SENSOR CHECK".B7_3.Memory_Bit_1,
           Memory_Bit_2             := "DB SENSOR CHECK".B7_3.Memory_Bit_2,
           Word_Buffer              := "DB SENSOR CHECK".B7_3.Word_buffer,
           Word_Result              := "DB SENSOR CHECK".B7_3.Word_Result);

NETWORK
TITLE =

